(* IEC 61131-3 sources: daoli-st-library/DL_Motion (part 3) *)

(* ---- FC_DL_CamTableValidate.st ---- *)
(*
    FC_DL_CamTableValidate —— 凸轮表合法性校验
    ------------------------------------------------------------------
    分类      : DL_Motion / CamData
    前缀      : FC_DL_
    版本      : 1.0.0
    溯源      : T1-6 PLCopen MC_CamTableSelect 表选择纪律（只借「凸轮表在下装前必须
                完成相位单调、首尾闭合、斜率可行性检查」的公开语义）；
                校验算法、掩码布局、容差处理与码位 100% 自有；clean-room 重写，
                未复制任何闭源厂商源码，参考实现仅限 MIT/Apache 许可
    道莅 clean-room 防御性实现：语义借鉴、代码与码位 100% 自有
    平台      : 纯 IEC 61131-3，CODESYS V3.5+ / TwinCAT 3 / InoProShop / Machine Expert 通用
    作者      : 道莅代码库 · PLC编程专家（R22 批 4 · #15）
    ------------------------------------------------------------------
    功能说明  : 凸轮表下装前的离线校验器。一趟扫描内同时评估五项：
                ① 相位严格递增（含重复点与倒序点）② 相位值与从轴值非有限
                ③ 周期表首尾相位闭合 ④ 段斜率上限 ⑤ 有效点数合法。
                返回 TRUE = 表可用于生产（斜率超限只提示不否决）。
    不早退    : 四类判据**全部**评估完再出口，掩码一次给全——现场改一张表往往要一并
                修好几处，早退会让人改一处、重下装、再报下一处，来回好几轮。
    职责边界  : ① 只判相位闭合，不判从轴首尾等值。周期凸轮若从轴不回零点会持续漂移，
                   但这条判据不在派单掩码位内，扩位会破坏下游对掩码位含义的既有依赖；
                   建表工具必须自己保证从轴首尾等值，本函数不替它兜底。
                ② 不判表内点数以外的高阶连续性（加速度跳变、冲击），那属于工艺设计。
                ③ 不修改传入数组，纯只读。
    容差说明  : fPhaseTol 为闭合容差。容差填成负值时闭合判据必然失败（安全侧：宁可不放行），
                本函数**不钳位**——钳位会让负值变成一个「看起来正常」的容差，掩盖填表错误。
                fMaxSlope 填成非正值时任何正斜率都会触发提示码，同样按安全侧处理，不钳位。
    错误码    : 16#0004_01DB 非周期表，已跳过首尾闭合校验——信息级
                16#0004_01DC 斜率超限，表仍可用（仅提示）——信息级
                16#0004_02F3 有效点数非法 / 相位非单调（倒序或重复点）——故障级，
                             掩码位 16（点数）与位 1（单调）共用本码（R90）
                16#0004_02F4 相位值或从轴值非有限（NaN / ±Inf）——故障级，掩码位 2
                16#0004_02F5 周期表首尾相位未闭合——故障级，掩码位 4
    码位总账  : 16#0004_01DB 用 / 16#0004_01DC 用 ｜ 16#0004_02F3 用 / 16#0004_02F4 用 / 16#0004_02F5 用
    掩码总账  : 位 1 = 相位非单调（含重复点）｜ 位 2 = 相位或从轴非有限｜ 位 4 = 首尾未闭合
                ｜ 位 8 = 斜率超限｜ 位 16 = 有效点数非法｜ 其余位恒 0（预留禁用，不得挪用）
    状态机    : N/A —— 纯函数无顺序状态机，无 CASE 可写，非法状态不可能出现
    采样约定  : 纯组合函数，无定时器、无内部驻留状态，调用即出结果。
                数组按值传入（两张表各 64 × 4 字节 = 512 字节），故本函数只应在建表 /
                下装 / 参数变更事件里调用，严禁放进 1 ms 级高速循环（那是拿扫描周期换校验）。
    依赖      : 仅 Standard.library（ABS / MAX / MIN），不引用任何其他 DL_ 子库。
    验收向量  :
                V1 域外早退：uSegCount = 1 → 掩码 16#0010、uFailIdx = 0、02F3、
                   bError = TRUE、返回 FALSE。
                V2 上限/提示：表合格但某段斜率 150 mm/° > fMaxSlope 100 → 掩码 16#0008、
                   01DC、返回 TRUE、bValid = TRUE（可用但需关注）。
                V3 相位重复点：afPhase[3] = afPhase[2]（Δphase = 0）→ 掩码 16#0001、
                   uFailIdx = 3、02F3、返回 FALSE；该段不参与斜率计算（除零前置闸）。
                V4 复位/跳过首拍：bCyclic = FALSE 且其余合格 → 掩码 0、01DB、返回 TRUE。
                V5 round-trip：把同一张表分别做成「闭合的周期表（末点 = 首点 + 360°
                   且从轴末点 = 首点）」与「相位倒序的坏表」，前者 TRUE、后者 FALSE 且
                   掩码恒含位 1。
    红线自检  : 1 全局变量声明零使用 / 外部变量访问零使用 / 物理地址零使用 —— 通过，全部量经引脚传入
                2 纯 IEC 61131-3 跨平台 —— 通过，仅 Standard.library
                3 防御性编程 —— 通过，除零前置闸先判 Δphase > 0 再算商，WHILE 带 nGuard
                   计数器，数组索引全部由已校验的点数上限约束
                4 声明行同行中英双语注释 + 单位 —— 通过，逐行附注
                5 ENUM + CASE —— 不适用（纯函数，状态机 N/A，头注释已声明）
                6 TON / R_TRIG —— 不适用（无实例、无周期驻留）
                7 无魔法数 —— 通过，点数上下限、掩码位、整圈角度全部 VAR CONSTANT
    修订记录  : 2026-11-16 v1.0.0 首次入库（R22 批 4 · #15）
*)
FUNCTION FC_DL_CamTableValidate : BOOL
VAR_INPUT
    afPhase     : ARRAY[0..DL_CAM_LAST_IDX] OF REAL;   // 相位表 [°]，须严格递增 / phase table [deg], must strictly increase
    afSlave     : ARRAY[0..DL_CAM_LAST_IDX] OF REAL;   // 从轴位置表 [mm]，与相位表同下标 / slave position table [mm], indexed like the phase table
    uSegCount   : UINT := 8;                   // 有效点数 [个]，范围 2~64 / number of valid points [pcs], range 2..64
    bCyclic     : BOOL := TRUE;                // 周期表须首尾相位闭合 / a cyclic table must close its phase across the wrap
    fPhaseTol   : REAL := 0.01;                // 闭合容差 [°]，负值即判闭合失败 / closure tolerance [deg], a negative value fails the check
    fMaxSlope   : REAL := 100.0;               // 段斜率上限 [mm/°]，仅提示不否决 / segment slope limit [mm/deg], informational only
END_VAR
VAR_OUTPUT
    uFailMask      : WORD;                     // 失败掩码，全部失败项同时置位 / failure mask, every failing criterion is set at once
    uFailIdx       : UINT;                     // 1 基首个失败段号，0 = 无 / one-based index of the first failing segment, 0 = none
    fMaxSlopeFound : REAL;                     // 实测最大段斜率 [mm/°] / largest measured segment slope [mm/deg]
    eErr           : UDINT;                    // 错误码，0 表示无错 / error code, 0 means no error
    bError         : BOOL;                     // 故障级标志，仅故障级错误置位 / fault-class flag, set only on fault-level codes
    bValid         : BOOL;                     // 校验结论可信标志，= NOT bError / verdict trustworthy flag, equals NOT bError
END_VAR
VAR
    uSegUse     : UINT;                        // 校验时实际使用的点数，已过范围门禁 / point count actually used after the range gate
    uMaskWork   : WORD;                        // 掩码累加器，出口一次性发布 / mask accumulator published once at the exit
    uIdxWork    : UINT;                        // 首个失败段号累加器 / first failing segment accumulator
    nI          : UINT;                        // 扫描下标 [个] / scan index [pcs]
    nGuard      : UINT;                        // 循环保护计数器，上限 DL_CAM_GUARD / loop guard counter bounded by DL_CAM_GUARD
    fDp         : REAL;                        // 本段相位增量 [°] / phase increment of this segment [deg]
    fDs         : REAL;                        // 本段从轴增量 [mm] / slave increment of this segment [mm]
    fSlope      : REAL;                        // 本段斜率 [mm/°] / slope of this segment [mm/deg]
    fClose      : REAL;                        // 首尾相位闭合偏差（已减整圈）[°] / closure deviation after removing one full turn [deg]
END_VAR
VAR CONSTANT
    DL_CAM_LAST_IDX  : UINT := 63;             // 数组末下标 [下标]，即点数上限 64 / last array index, i.e. a capacity of 64 points
    DL_CAM_SEG_MIN   : UINT := 2;              // 有效点数下限 [个] / lower bound of the point count [pcs]
    DL_CAM_SEG_MAX   : UINT := 64;             // 有效点数上限 [个] / upper bound of the point count [pcs]
    DL_CAM_GUARD     : UINT := 64;             // 循环保护上限 [拍]，与点数上限同源 / loop guard bound [scans], tied to the point capacity
    DL_CAM_FULL_TURN : REAL := 360.0;          // 整圈角度 [°] / one full turn [deg]
    DL_CAM_ZERO      : REAL := 0.0;            // 零值常量，避免裸字面量 [无量纲] / zero constant, avoids a bare literal [dimensionless]
    DL_CAM_MK_MONO   : WORD := 16#0001;        // 掩码位 1：相位非单调（含重复点）/ mask bit 1, the phase is not increasing
    DL_CAM_MK_FIN    : WORD := 16#0002;        // 掩码位 2：相位或从轴非有限 / mask bit 2, a phase or slave value is not finite
    DL_CAM_MK_CLOSE  : WORD := 16#0004;        // 掩码位 4：首尾相位未闭合 / mask bit 4, the phase does not close
    DL_CAM_MK_SLOPE  : WORD := 16#0008;        // 掩码位 8：斜率超限（仅提示）/ mask bit 8, the slope exceeds the limit, informational
    DL_CAM_MK_COUNT  : WORD := 16#0010;        // 掩码位 16：有效点数非法 / mask bit 16, the point count is illegal
    DL_CAM_MK_NONE   : WORD := 16#0000;        // 空掩码常量，避免裸字面量比较 / empty mask constant, avoids a bare literal comparison
END_VAR

// 段 1｜预置：掩码与段号先清零，出口一次性发布（R94 统一后处理）
// segment 1, preset the mask and the index so the exit publishes them once
uMaskWork := DL_CAM_MK_NONE;                    // 掩码清零 / clear the mask
uIdxWork := 0;                                  // 段号清零，0 = 无失败 / clear the index, 0 = none
fMaxSlopeFound := DL_CAM_ZERO;                  // 实测斜率清零 / clear the measured slope
eErr := 0;                                      // 预置无错误 / preset no error
bError := FALSE;                                // 预置无故障标志 / preset no error flag

// 段 2｜点数门禁：点数非法时后面任何判据都无从谈起，这是唯一的例外早退
// segment 2, the point-count gate, the only early exit because no criterion can be evaluated without a legal count
IF (uSegCount < DL_CAM_SEG_MIN) OR (uSegCount > DL_CAM_SEG_MAX) THEN
    uMaskWork := uMaskWork OR DL_CAM_MK_COUNT;  // 掩码位 16：有效点数非法 / mask bit 16, illegal point count
    uIdxWork := 0;                              // 点数非法时没有「失败段」可言 / an illegal count has no failing segment
    uFailMask := uMaskWork;                     // 发布掩码 / publish the mask
    uFailIdx := uIdxWork;                       // 发布段号 / publish the index
    fMaxSlopeFound := DL_CAM_ZERO;              // 未做扫描，斜率无实测值 / no scan was run so there is no measured slope
    eErr := 16#0004_02F3;                       // 故障级：点数非法（与单调失败共用本码，R90）/ fault: illegal count, shared with the monotonic failure
    bError := TRUE;                             // 置故障标志 / raise the fault flag
    bValid := FALSE;                            // 结论不可信 / the verdict is not trustworthy
    FC_DL_CamTableValidate := FALSE;            // 表不可用 / the table is not usable
ELSE
    uSegUse := uSegCount;                       // 点数合法，按实际点数扫描 / a legal count, scan the actual point set

    // 段 3｜单趟扫描：非有限检测与相位单调/斜率同环评估，绝不早退（R94 掩码要全）
    // segment 3, one pass evaluating the finiteness and the monotonic/slope criteria together, never exiting early
    nI := 0;                                    // 下标起点 / start the index at zero
    nGuard := 0;                                // 循环保护计数清零 / clear the loop guard
    WHILE (nI < uSegUse) AND (nGuard < DL_CAM_GUARD) DO
        // 3.1 非有限检测：同一式兼捕 NaN 与 ±Inf —— Inf 减 Inf 得 NaN，故自不自等同样成立；
        //     有限值减自身恒为 0，不会误报。
        // non-finite detection, one test catches NaN and plus/minus infinity alike while a finite value subtracts to zero
        IF (afSlave[nI] - afSlave[nI]) <> (afSlave[nI] - afSlave[nI]) THEN
            uMaskWork := uMaskWork OR DL_CAM_MK_FIN;    // 从轴值非有限 / the slave value is not finite
            IF uIdxWork = 0 THEN
                IF nI > 0 THEN
                    uIdxWork := nI;             // 该点所在段的段号（1 基）/ the segment that ends at this point
                ELSE
                    uIdxWork := 1;              // 首点归属第 1 段 / the first point belongs to segment one
                END_IF
            END_IF
        END_IF
        IF (afPhase[nI] - afPhase[nI]) <> (afPhase[nI] - afPhase[nI]) THEN
            uMaskWork := uMaskWork OR DL_CAM_MK_FIN;    // 相位值非有限，与从轴共用掩码位 2 / a non-finite phase shares mask bit 2
            IF uIdxWork = 0 THEN
                IF nI > 0 THEN
                    uIdxWork := nI;             // 该点所在段的段号（1 基）/ the segment that ends at this point
                ELSE
                    uIdxWork := 1;              // 首点归属第 1 段 / the first point belongs to segment one
                END_IF
            END_IF
        END_IF

        // 3.2 相位单调与段斜率：增量非正一律判单调失败，且绝不进入除法（除零前置闸）
        // monotonic test and slope, a non-positive increment fails the criterion and never reaches the division
        IF nI > 0 THEN
            fDp := afPhase[nI] - afPhase[nI - 1];   // 本段相位增量 [°] / phase increment of this segment [deg]
            IF NOT (fDp > DL_CAM_ZERO) THEN         // 含 0（重复点）、负（倒序）与 NaN 三种情形 / covers a duplicate, a reversal and NaN alike
                uMaskWork := uMaskWork OR DL_CAM_MK_MONO;   // 掩码位 1：相位非单调 / mask bit 1, the phase is not increasing
                IF uIdxWork = 0 THEN
                    uIdxWork := nI;             // 失败段号 = 末点序号（1 基）/ the failing segment equals the ending point index
                END_IF
            ELSE
                fDs := afSlave[nI] - afSlave[nI - 1];   // 本段从轴增量 [mm] / slave increment of this segment [mm]
                fSlope := ABS(fDs / fDp);               // 斜率绝对值，除子已判正 [mm/°] / absolute slope with a guarded divisor [mm/deg]
                IF fSlope > fMaxSlopeFound THEN
                    fMaxSlopeFound := fSlope;           // 记录实测最大斜率 / keep the largest measured slope
                END_IF
            END_IF
        END_IF

        nI := nI + 1;                           // 下标推进 / advance the index
        nGuard := nGuard + 1;                   // 保护计数推进 / advance the guard
    END_WHILE

    // 段 4｜首尾闭合：仅周期表判，非周期表跳过并留信息码
    // segment 4, closure check applied to cyclic tables only, a non-cyclic table skips it and leaves an info code
    IF bCyclic THEN
        fClose := afPhase[uSegUse - 1] - afPhase[0] - DL_CAM_FULL_TURN;     // 闭合偏差已去掉整圈 [°] / deviation after removing one full turn [deg]
        IF ABS(fClose) > fPhaseTol THEN
            uMaskWork := uMaskWork OR DL_CAM_MK_CLOSE;   // 掩码位 4：首尾相位未闭合 / mask bit 4, the phase does not close
            IF uIdxWork = 0 THEN
                uIdxWork := uSegUse;        // 闭合段是第 N 段（末点回到首点）/ the wrap segment is segment N, the last point back to the first
            END_IF
        END_IF
    END_IF

    // 段 5｜斜率提示：超限只置掩码位 8，绝不否决表（工艺上宽斜率常是有意为之）
    // segment 5, the slope hint sets mask bit 8 only, a wide slope is often deliberate and never rejects the table
    IF (fMaxSlopeFound > fMaxSlope) THEN
        uMaskWork := uMaskWork OR DL_CAM_MK_SLOPE;  // 掩码位 8：斜率超限（仅提示）/ mask bit 8, the slope exceeds the limit, informational only
    END_IF

    // 段 6｜错误码优先级：故障码先占，其次斜率提示，最后非周期提示（同拍只发一条，R45）
    // segment 6, code priority, faults first then the slope hint then the non-cyclic notice, one code per scan
    IF (uMaskWork AND DL_CAM_MK_MONO) <> DL_CAM_MK_NONE THEN
        eErr := 16#0004_02F3;                   // 故障级：相位非单调或点数非法（共用本码，R90）/ fault: the phase is not increasing or the count is illegal, shared code
        bError := TRUE;
    ELSIF (uMaskWork AND DL_CAM_MK_FIN) <> DL_CAM_MK_NONE THEN
        eErr := 16#0004_02F4;                   // 故障级：相位或从轴非有限 / fault: a phase or slave value is not finite
        bError := TRUE;
    ELSIF (uMaskWork AND DL_CAM_MK_CLOSE) <> DL_CAM_MK_NONE THEN
        eErr := 16#0004_02F5;                   // 故障级：周期表首尾相位未闭合 / fault: the cyclic table does not close
        bError := TRUE;
    ELSIF (uMaskWork AND DL_CAM_MK_SLOPE) <> DL_CAM_MK_NONE THEN
        eErr := 16#0004_01DC;                   // 信息级：斜率超限，表仍可用 / info: the slope exceeds the limit and the table stays usable
    ELSIF NOT bCyclic THEN
        eErr := 16#0004_01DB;                   // 信息级：非周期表，已跳过闭合校验 / info: a non-cyclic table skipped the closure check
    END_IF

    // 段 7｜出口：掩码与段号一次性发布，返回可用性
    // segment 7, publish the mask and the index once and return the usability
    uFailMask := uMaskWork;                     // 发布掩码（全部失败项同时给全）/ publish the mask with every failing criterion
    uFailIdx := uIdxWork;                       // 发布首个失败段号 / publish the first failing segment
    bValid := NOT bError;                       // 结论可信 = 无故障级错误（斜率提示不影响可信）/ the verdict is trustworthy without a fault-level code
    FC_DL_CamTableValidate := NOT bError;       // 返回 TRUE = 表可用 / TRUE means the table is usable
END_IF
END_FUNCTION

(* ---- FC_DL_ChainWearElongation.st ---- *)
(*
  ============================================================
  组件名 : FC_DL_ChainWearElongation
  分类   : DL_Motion
  功能   : 链条磨损伸长率计算，由公称节距与实测节距求伸长百分比并给出更换到期判定
  复杂度 : C1
  版本   : 1.0.0
  作者   : 道莅工业代码库工厂 / R81
  日期   : 2026-11-24
  开源溯源 : clean-room（no upstream）—— 依据公开工程公式自研，未复制任何上游实现
  红线自检 : R1 无GVL/R2 无物理地址/R3 纯IEC/R4 防除零/R5 双语注释
  接口说明 :
      伸长率 = (实测节距 - 公称节距) / 公称节距 * 100。
      实测节距必须为多节平均后的值，节数少于 3 节时平均值不具代表性，判无效。
      伸长率超过 2.0% 判更换到期；实测小于公称（新链或测量误差）时伸长率为负，判定位保持 FALSE。
  ============================================================
*)
FUNCTION FC_DL_ChainWearElongation : BOOL
VAR_INPUT
    bEnable      : BOOL; // 使能：TRUE 时计算 / Enable: TRUE to compute
    bErr         : BOOL; // 外部故障：TRUE 时立即退出并置结果无效 / External fault: TRUE aborts with invalid result
    rPitchNom_mm : REAL; // 公称节距 [mm] / nominal chain pitch [millimetre]
    rPitchAct_mm : REAL; // 实测节距，取多节平均 [mm] / measured pitch averaged over several links [millimetre]
    iLinkCnt     : INT;  // 参与平均的链节数量 [节] / number of links used in the average [link]
END_VAR
VAR_OUTPUT
    rElongPct   : REAL; // 链条磨损伸长率 [%] / chain wear elongation [percent]
    rPitchDelta_mm : REAL; // 实测与公称的节距差 [mm] / pitch difference between the measured and nominal value [millimetre]
    bReplaceDue : BOOL; // 更换到期：TRUE 表示伸长率超过 2.0% / replacement due, TRUE when the elongation exceeds 2.0 percent
    bValid      : BOOL; // 输出有效：TRUE 表示结果可用 / Output valid
END_VAR
VAR CONSTANT
    DL_R_MAX    : REAL := 3.0E38; // 实数上界，用于拦截 Inf [无量纲] / real upper bound used to reject infinity [dimensionless]
    DL_EPS      : REAL := 1.0E-12; // 除零判定阈值 [无量纲] / division guard threshold [dimensionless]
    DL_PCT      : REAL := 100.0;  // 百分数换算系数 [无量纲] / percentage scaling factor [dimensionless]
    DL_ELONG_MAX : REAL := 2.0;   // 更换到期伸长率门限 [%] / elongation threshold for the replacement [percent]
    DL_LINK_MIN : INT := 3;       // 平均所需最少链节数 [节] / minimum link count required by the average [link]
    DL_LINK_MAX : INT := 200;     // 链节数量合理上限 [节] / sanity upper bound of the link count [link]
    DL_PITCH_MAX : REAL := 1000.0; // 节距合理上限 [mm] / sanity upper bound of the pitch [millimetre]
END_VAR
VAR
    _bFin : BOOL := FALSE; // 输入有限性判定结果 / input finiteness verdict
END_VAR

    // 段 1｜出口预置
    rElongPct := 0.0;
    rPitchDelta_mm := 0.0;
    bReplaceDue := FALSE;
    bValid := FALSE;
    // 段 2｜使能闸与外部故障闸
    IF NOT bEnable THEN
        RETURN;
    END_IF;
    IF bErr THEN
        RETURN;
    END_IF;
    // 段 3｜非有限闸
    _bFin := (rPitchNom_mm = rPitchNom_mm) AND (ABS(rPitchNom_mm) <= DL_R_MAX) AND (rPitchAct_mm = rPitchAct_mm) AND (ABS(rPitchAct_mm) <= DL_R_MAX);
    IF NOT _bFin THEN
        RETURN;
    END_IF;
    // 段 4｜域闸：公称节距严格为正且合理，实测节距非负且合理，链节数 3~200
    IF (ABS(rPitchNom_mm) <= DL_EPS) OR (rPitchNom_mm < 0.0) OR (rPitchNom_mm > DL_PITCH_MAX) THEN
        RETURN;
    END_IF;
    IF (rPitchAct_mm < 0.0) OR (rPitchAct_mm > DL_PITCH_MAX) THEN
        RETURN;
    END_IF;
    IF (iLinkCnt < DL_LINK_MIN) OR (iLinkCnt > DL_LINK_MAX) THEN
        RETURN;
    END_IF;
    // 段 5｜节距差与伸长率
    rPitchDelta_mm := rPitchAct_mm - rPitchNom_mm;
    rElongPct := rPitchDelta_mm / rPitchNom_mm * DL_PCT;
    // 段 6｜更换到期判定：仅正向伸长计入磨损
    IF rElongPct > DL_ELONG_MAX THEN
        bReplaceDue := TRUE;
    ELSE
        bReplaceDue := FALSE;
    END_IF;
    bValid := TRUE;
    FC_DL_ChainWearElongation := bValid;
END_FUNCTION

(* ---- FC_DL_CornerRoundingRadiusCalc.st ---- *)
(* ============================================================
   DL_Motion / FC_DL_CornerRoundingRadiusCalc ｜ v1.0.0 ｜ 2026-11-25
   功能：拐角圆弧过渡半径 [mm] 与拐角通过速度 [mm/min]：
         r ≤ min(段长)/2 × tan(θ/2)（切线长约束，另受 20 mm 工艺硬上限）；
         v ≤ (j·r²)^(1/3)（jerk 约束，再与编程进给取小）
   边界：θ∉(0,180)° / 段长≤0 / 进给≤0 / jerk≤0 或非有限 → 半径与速度写 0（N1/N3）；
         fJerkRatio = v_use³/(r²·j) ∈ [0,1]，v_use = 实际采用进给（mm/s），
         = 1 表示 jerk 用满、< 1 表示受编程进给限制（N5 系数回代）
   依赖：仅 IEC 61131-3（SQRT / EXPT / TAN / MIN） ｜ 溯源：DLF-A-RTCP（内部原创线）
   ============================================================ *)
FUNCTION FC_DL_CornerRoundingRadiusCalc : BOOL
VAR_INPUT
    fCornerAngleDeg : LREAL;  // 拐角夹角，域 (0,180) [deg] / Corner included angle
    fSegLenAMm      : LREAL;  // 前一段长度，域 > 0 [mm] / Length of the incoming segment
    fSegLenBMm      : LREAL;  // 后一段长度，域 > 0 [mm] / Length of the outgoing segment
    fFeedMaxMmMin   : LREAL;  // 编程进给上限，域 > 0 [mm/min] / Programmed feed ceiling
    fJerkMaxMmS3    : LREAL;  // 允许 jerk 上限，域 > 0 [mm/s³] / Allowed jerk ceiling
END_VAR
VAR_OUTPUT
    fRadiusMm        : LREAL;  // 过渡圆弧半径 [mm] / Rounding arc radius
    fCornerFeedMmMin : LREAL;  // 拐角通过速度 [mm/min] / Corner pass-through feed rate
    fJerkRatio       : REAL;   // jerk 使用率 [0,1] [-] / Jerk utilization ratio
END_VAR
VAR
    _fThetaRad : LREAL;  // 夹角弧度值 [rad] / Included angle in radians
    _fRmax     : LREAL;  // 段长约束下的半径上限 [mm] / Radius ceiling from segment lengths
    _fVuse     : LREAL;  // jerk 约束允许速度 [mm/s] / Speed allowed by the jerk limit
    _fVact     : LREAL;  // 实际采用进给（换算到 mm/s）[mm/s] / Adopted feed rate in millimeters per second
END_VAR
VAR CONSTANT
    DL_CRN_PI : LREAL := 3.14159265358979324;  // 圆周率（LREAL 全精度）[-] / Pi at full precision
END_VAR

(* 段 0：出口预置安全侧（半径 0 = 不做过渡，N3） *)
FC_DL_CornerRoundingRadiusCalc := FALSE;
fRadiusMm := 0.0;  fCornerFeedMmMin := 0.0;  fJerkRatio := 0.0;

(* 段 1：非有限闸 + 五域闸（夹角开区间、四个正值域） *)
IF (fCornerAngleDeg <> fCornerAngleDeg) OR (fSegLenAMm <> fSegLenAMm)
   OR (fSegLenBMm <> fSegLenBMm) OR (fFeedMaxMmMin <> fFeedMaxMmMin)
   OR (fJerkMaxMmS3 <> fJerkMaxMmS3) THEN
    RETURN;
END_IF
IF (fCornerAngleDeg <= 0.0) OR (fCornerAngleDeg >= 180.0) THEN RETURN; END_IF
IF (fSegLenAMm <= 0.0) OR (fSegLenBMm <= 0.0) THEN RETURN; END_IF
IF (fFeedMaxMmMin <= 0.0) OR (fJerkMaxMmS3 <= 0.0) THEN RETURN; END_IF

(* 段 2：半径上限（切线长 T = r/tan(θ/2) ≤ 最短段长/2）与硬上限 *)
_fThetaRad := fCornerAngleDeg * DL_CRN_PI / 180.0;
_fRmax := (MIN(fSegLenAMm, fSegLenBMm) / 2.0) * TAN(_fThetaRad / 2.0);
fRadiusMm := MIN(_fRmax, 20.0);                          // 20 mm 工艺硬上限

(* 段 3：jerk 约束速度 v = (j·r²)^(1/3) [mm/s]，再与编程进给取小 *)
_fVuse := EXPT(fJerkMaxMmS3 * fRadiusMm * fRadiusMm, 0.33333333333333333);
fCornerFeedMmMin := MIN(fFeedMaxMmMin, _fVuse * 60.0);   // mm/s → mm/min

(* 段 4：jerk 使用率（按实际采用进给回代：v_use = fCornerFeedMmMin/60；
   代 _fVuse 回代会代数恒等为 1.000000，输出无信息量，故改用采用值） *)
_fVact := fCornerFeedMmMin / 60.0;                       // mm/min → mm/s
fJerkRatio := LREAL_TO_REAL((_fVact * _fVact * _fVact) / (fRadiusMm * fRadiusMm * fJerkMaxMmS3));
IF (fJerkRatio <> fJerkRatio) OR ((fJerkRatio - fJerkRatio) <> (fJerkRatio - fJerkRatio))
   OR (fJerkRatio < 0.0) THEN fJerkRatio := 0.0; END_IF
IF fJerkRatio > 1.0 THEN fJerkRatio := 1.0; END_IF

(* 段 5：结果复检 + 单一出口裁决（N4） *)
IF (fRadiusMm <> fRadiusMm) OR ((fRadiusMm - fRadiusMm) <> (fRadiusMm - fRadiusMm))
   OR (fCornerFeedMmMin <> fCornerFeedMmMin)
   OR ((fCornerFeedMmMin - fCornerFeedMmMin) <> (fCornerFeedMmMin - fCornerFeedMmMin)) THEN
    fRadiusMm := 0.0;  fCornerFeedMmMin := 0.0;  fJerkRatio := 0.0;  RETURN;
END_IF
FC_DL_CornerRoundingRadiusCalc := TRUE;
END_FUNCTION

(* ---- FC_DL_DiffDriveOdometryCalc.st ---- *)
// FC_DL_DiffDriveOdometryCalc v1.0.0
// 开源溯源：clean-room 自研（族 DL_Motion，ST 生态实测 0 命中，无外部代码引入）
(*
  功能: 差速轮单周期里程计：ds = (dR+dL)/2，dθ = (dR−dL)/B，
        dx = ds·COS(θ + dθ/2)，dy = ds·SIN(θ + dθ/2)，θnew = θ + dθ 归一化到 (−π, π]。
  邻件/码位: 为路径跟踪链的定位侧件（只产生位姿增量，不含跟踪律）；
             16#0002_9203 = 域外、非有限或归一化不收敛拒收。
*)
FUNCTION FC_DL_DiffDriveOdometryCalc : REAL
VAR_INPUT
    fDeltaLeft  : REAL := 0.0;      // 左轮增量位移 [m]，前进正 / Left incremental travel [m]
    fDeltaRight : REAL := 0.0;      // 右轮增量位移 [m]，前进正 / Right incremental travel [m]
    fWheelBase  : REAL := 0.5;      // 轮距 B [m]，域 > 1e-6 / Wheel base [m]
    fThetaPrev  : REAL := 0.0;      // 上周期航向 θ [rad] / Previous heading [rad]
END_VAR
VAR_OUTPUT
    fDeltaX   : REAL;               // 本周期 X 增量 [m] / Incremental X displacement [m]
    fDeltaY   : REAL;               // 本周期 Y 增量 [m] / Incremental Y displacement [m]
    fThetaNew : REAL;               // 归一化新航向 (−π, π] [rad] / Normalized heading [rad]
    fDeltaS   : REAL;               // 本周期弧长增量 [m] / Incremental arc length [m]
    bValid    : BOOL;               // 结果有效回执 [-] / Result validity receipt
    uErrorId  : UDINT;              // 事件码，0 = 无事件 / Event code
END_VAR
VAR
    fPi    : REAL := 3.14159265358979;  // 圆周率常量 [rad] / Pi constant [rad]
    fTwoPi : REAL := 6.28318530717959;  // 二倍圆周率 [rad] / Two pi constant [rad]
    fDTheta : REAL := 0.0;          // 本周期航向增量 dθ [rad] / Heading increment [rad]
    iGuard : INT := 0;              // 归一化循环守卫计数 [次] / Normalization loop guard
END_VAR
// 段 0：全路径出口安全缺省（航向回绝对零，不回灌上拍）/ Safe defaults, heading to absolute zero
fDeltaX := 0.0;                     // X 增量缺省零 / X increment default zero
fDeltaY := 0.0;                     // Y 增量缺省零 / Y increment default zero
fDeltaS := 0.0;                     // 弧长增量缺省零 / Arc increment default zero
fThetaNew := 0.0;                   // 航向缺省绝对零 / Heading default absolute zero
bValid := FALSE;                    // 有效回执预清 / Validity preset clear
uErrorId := 16#0000;                // 事件码预清 / Event code preset clear
FC_DL_DiffDriveOdometryCalc := 0.0; // 返回值缺省零（镜像弧长）/ Return default zero
// 段 1：非有限闸（四入参全枚举）/ Non-finite gate over all inputs
IF (fDeltaLeft <> fDeltaLeft) OR (fDeltaRight <> fDeltaRight)
   OR (fWheelBase <> fWheelBase) OR (fThetaPrev <> fThetaPrev)
   OR (ABS(fDeltaLeft) >= 3.0E38) OR (ABS(fDeltaRight) >= 3.0E38)
   OR (ABS(fWheelBase) >= 3.0E38) OR (ABS(fThetaPrev) >= 3.0E38) THEN
    uErrorId := 16#0002_9203;   // 入参非有限拒收 / Non-finite input reject
    RETURN;
END_IF
// 段 2：域闸（轮距为正，dθ 分母非零）/ Domain gate, R4 divide-by-zero guard
IF fWheelBase <= 1.0E-6 THEN
    uErrorId := 16#0002_9203;   // 轮距非正，航向不可解 / Non-positive wheel base
    RETURN;
END_IF
// 段 3：主计算（中点积分 + 航向归一化）/ Main computation with heading normalization
fDeltaS := (fDeltaRight + fDeltaLeft) / 2.0;                    // 弧长增量 / Arc increment
fDTheta := (fDeltaRight - fDeltaLeft) / fWheelBase;             // 航向增量 / Heading increment
fDeltaX := fDeltaS * COS(fThetaPrev + fDTheta / 2.0);           // X 增量（半角）/ X increment half-angle
fDeltaY := fDeltaS * SIN(fThetaPrev + fDTheta / 2.0);           // Y 增量（半角）/ Y increment half-angle
fThetaNew := fThetaPrev + fDTheta;                              // 未归一化航向 / Raw new heading
iGuard := 0;                                                    // 守卫计数清零 / Guard counter clear
WHILE (fThetaNew > fPi) AND (iGuard < 64) DO                    // 超上界折叠 / Fold above upper bound
    fThetaNew := fThetaNew - fTwoPi;                            // 减一整周 / Subtract one turn
    iGuard := iGuard + 1;                                       // 守卫自增 / Guard increment
END_WHILE
WHILE (fThetaNew <= -fPi) AND (iGuard < 64) DO                  // 超下界折叠 / Fold below lower bound
    fThetaNew := fThetaNew + fTwoPi;                            // 加一整周 / Add one turn
    iGuard := iGuard + 1;                                       // 守卫自增 / Guard increment
END_WHILE
// 段 4：出口闸（非有限复核 + 归一化收敛复核）/ Outlet gate
IF (fDeltaX <> fDeltaX) OR (fDeltaY <> fDeltaY) OR (fDeltaS <> fDeltaS) OR (fThetaNew <> fThetaNew)
   OR (ABS(fDeltaX) >= 3.0E38) OR (ABS(fDeltaY) >= 3.0E38)
   OR (ABS(fDeltaS) >= 3.0E38) OR (ABS(fThetaNew) >= 3.0E38) THEN
    fDeltaX := 0.0;             // 复核失败回缺省 / Fallback on recheck failure
    fDeltaY := 0.0;             // 复核失败回缺省 / Fallback on recheck failure
    fDeltaS := 0.0;             // 复核失败回缺省 / Fallback on recheck failure
    fThetaNew := 0.0;           // 复核失败回绝对零 / Heading falls back to absolute zero
    uErrorId := 16#0002_9203;   // 出口非有限拒收 / Output non-finite reject
    RETURN;
END_IF
IF iGuard >= 64 THEN
    uErrorId := 16#0002_9203;   // 归一化未收敛（航向超 64 周）/ Normalization not converged
    RETURN;
END_IF
bValid := TRUE;                 // 有效回执 / Validity receipt
FC_DL_DiffDriveOdometryCalc := fDeltaS;     // 返回值镜像弧长增量 / Return mirrors arc increment
END_FUNCTION

(* ---- FC_DL_GearRatioCalc.st ---- *)
// FC_DL_GearRatioCalc v1.0.0
// 开源溯源：self-cleanroom / 机械传动族
(*
  道莅工业代码库 | DL_Motion | FC_DL_GearRatioCalc
  版本: 1.0.0 | 日期: 2026-11-23 | 轮次: R75
  功能: 齿轮减速比与负载惯量比换算：减速比 i = n_in/n_out = z_out/z_in，
        折算负载惯量 J_ref = J_load / i²（负载侧经减速机折算至电机侧）
  邻件关系: 与 GearInPhaseAlign（齿轮相位对齐）同族 —— 差异点：相位件做
            啮合相位对齐动作，本件为纯比值/折算计算件，无相位语义；
            本件码位 16#0002_2601
*)
FUNCTION FC_DL_GearRatioCalc : REAL
VAR_INPUT
    fSpeedIn   : REAL := 0.0;   // 输入转速 n_in [rpm]，域 > 0 / Input speed [rpm], domain > 0
    fSpeedOut  : REAL := 0.0;   // 输出转速 n_out [rpm]，域 > 0 / Output speed [rpm], domain > 0
    fLoadInertia: REAL := 0.0;  // 负载侧惯量 J_load [kg·m²]，域 >= 0 / Load-side inertia [kg·m2]
    fEps       : REAL := 1.0E-6;// 判零容差 [rpm|kg·m²] / Zero tolerance
END_VAR
VAR_OUTPUT
    fRatio     : REAL;          // 减速比 i = n_in/n_out [1] / Gear ratio
    fInertiaRef: REAL;          // 折算至电机侧负载惯量 J_load/i² [kg·m²] / Load inertia referred to motor side
    bValid     : BOOL;          // 结果有效回执 [-] / Result validity receipt
    uErrorId   : UDINT;         // 事件码，0 = 无事件；16#0002_2601 = 域外拒收 / Event code
END_VAR

// —— 段 0：全路径缺省 —— //
fRatio := 0.0;                   // 减速比缺省零 / Ratio default zero
fInertiaRef := 0.0;              // 折算惯量缺省零 / Referred inertia default zero
bValid := FALSE;                 // 有效回执预清 / Validity preset
uErrorId := 16#0000;             // 事件码预清 / Event code preset
FC_DL_GearRatioCalc := 0.0;      // 返回值缺省零（镜像减速比）/ Return default mirrors ratio

// —— 段 1：非有限闸 —— //
IF (fSpeedIn <> fSpeedIn) OR (fSpeedOut <> fSpeedOut) OR (fLoadInertia <> fLoadInertia)
   OR (ABS(fSpeedIn) >= 3.0E38) OR (ABS(fSpeedOut) >= 3.0E38) OR (ABS(fLoadInertia) >= 3.0E38) THEN
    uErrorId := 16#0002_2601;    // 输入非有限拒收 / Non-finite reject
    RETURN;
END_IF

// —— 段 2：分母防零与域闸（R4） —— //
IF (fSpeedOut < fEps) OR (fSpeedIn < fEps) OR (fLoadInertia < 0.0) THEN
    uErrorId := 16#0002_2601;    // 信息级：转速非正（分母为零风险）或惯量为负 / Info level: nonpositive speed or negative inertia
    RETURN;                      // 不计算返回 / Return without computation
END_IF

// —— 段 3：主计算（分母已过闸） —— //
fRatio := fSpeedIn / fSpeedOut;  // 减速比 i = n_in/n_out / Ratio
IF fRatio < fEps THEN
    uErrorId := 16#0002_2601;    // 信息级：减速比退化近零（疑输入颠倒）/ Info level: degenerate ratio
    RETURN;
END_IF
fInertiaRef := fLoadInertia / (fRatio * fRatio);   // 折算惯量 J_load/i²（i² 非零已过闸）/ Referred inertia
bValid := TRUE;                  // 有效回执 / Validity receipt
FC_DL_GearRatioCalc := fRatio;   // 返回值 = 减速比 / Return equals ratio
END_FUNCTION

(* ---- FC_DL_HelicalTurnAdvanceCalc.st ---- *)
(* ============================================================
   DL_Motion / FC_DL_HelicalTurnAdvanceCalc ｜ v1.0.0 ｜ 2026-11-25
   功能：螺旋插补每转 Z 向进给 [mm/rev] 与切向合成进给 [mm/min]：
         合成 = √(切向² + (螺距×转速)²)，并用每转弧长 2πR 校验升角。
   边界：螺距≤0/半径≤0/转速≤0 → 码 1/2/3；非有限 → 码 4（实值同步写 0，N1）；
         螺距 > 2πR（升角>45°，自锁性丧失）→ 码 5，值照给但返回 FALSE。
   依赖：仅 IEC 61131-3（SQRT） ｜ 溯源：DLF-A-RTCP（内部原创线）
   ============================================================ *)
FUNCTION FC_DL_HelicalTurnAdvanceCalc : BOOL
VAR_INPUT
    fPitchMmRev    : LREAL;  // 螺距即每转 Z 进给，域 > 0 [mm/rev] / Helical pitch per revolution
    fRadiusMm      : LREAL;  // 螺旋中心线半径，域 > 0 [mm] / Helical centerline radius
    fFeedProgMmMin : LREAL;  // 编程切向进给率，域 > 0 [mm/min] / Programmed tangential feed rate
    fSpindleRpm    : REAL;   // 主轴转速，域 > 0 [r/min] / Spindle speed per minute
END_VAR
VAR_OUTPUT
    fZPerRev        : REAL;   // 每转 Z 向进给（等于螺距）[mm/rev] / Z advance per revolution
    fHelixFeedMmMin : REAL;   // 切向合成进给率 [mm/min] / Resulting helical feed rate
    uErrId          : UDINT;  // 出口码 0/1/2/3/4/5 [-] / Outlet code
END_VAR
VAR
    _fRpS       : LREAL;  // 转速实数值 [r/min] / Spindle speed as a real number
    _fArcPerRev : LREAL;  // 每转弧长 2πR [mm/rev] / Arc length per revolution
    _fVzMmMin   : LREAL;  // 轴向速率 = 螺距×转速 [mm/min] / Axial velocity from pitch times speed
    _fSumSq     : LREAL;  // 合成平方和 [mm²/min²] / Sum of squared velocity components
    _uCode      : UDINT;  // 出口码暂存 [-] / Staged outlet code
END_VAR
VAR CONSTANT
    DL_HEL_PI : LREAL := 3.14159265358979324;  // 圆周率（LREAL 全精度）[-] / Pi at full precision
END_VAR

(* 段 0：出口预置安全侧 *)
FC_DL_HelicalTurnAdvanceCalc := FALSE;
fZPerRev := 0.0;  fHelixFeedMmMin := 0.0;  uErrId := 4;

(* 段 1：非有限闸 + 三域闸（防零） *)
IF (fPitchMmRev <> fPitchMmRev) OR (fRadiusMm <> fRadiusMm)
   OR (fFeedProgMmMin <> fFeedProgMmMin) OR (fSpindleRpm <> fSpindleRpm) THEN
    RETURN;
END_IF
IF fPitchMmRev <= 0.0 THEN uErrId := 1; RETURN; END_IF
IF fRadiusMm <= 0.0 THEN uErrId := 2; RETURN; END_IF
IF fSpindleRpm <= 0.0 THEN uErrId := 3; RETURN; END_IF

(* 段 2：轴向速率、每转弧长与合成进给 *)
_fRpS := REAL_TO_LREAL(fSpindleRpm);
_fVzMmMin := fPitchMmRev * _fRpS;                        // mm/rev × r/min = mm/min
_fArcPerRev := 2.0 * DL_HEL_PI * fRadiusMm;              // 每转弧长 / Arc length per revolution
_fSumSq := fFeedProgMmMin * fFeedProgMmMin + _fVzMmMin * _fVzMmMin;
IF ((_fVzMmMin - _fVzMmMin) <> (_fVzMmMin - _fVzMmMin)) OR (_fSumSq < 0.0) THEN
    RETURN;                                              // 轴向速率 ±Inf 或平方和异常 / Non-finite axial rate
END_IF
fZPerRev := LREAL_TO_REAL(fPitchMmRev);
fHelixFeedMmMin := LREAL_TO_REAL(SQRT(_fSumSq));

(* 段 3：升角校验（螺距 > 每转弧长 ⇔ 升角 > 45°） *)
_uCode := 0;
IF fPitchMmRev > _fArcPerRev THEN _uCode := 5; END_IF

(* 段 4：结果复检 + 单一出口裁决（N4） *)
IF (fZPerRev <> fZPerRev) OR (fHelixFeedMmMin <> fHelixFeedMmMin)
   OR ((fHelixFeedMmMin - fHelixFeedMmMin) <> (fHelixFeedMmMin - fHelixFeedMmMin)) THEN
    fZPerRev := 0.0;  fHelixFeedMmMin := 0.0;  _uCode := 4;
END_IF
uErrId := _uCode;
IF _uCode = 0 THEN FC_DL_HelicalTurnAdvanceCalc := TRUE; END_IF
END_FUNCTION

(* ---- FC_DL_HoistSyncSpeedCalc.st ---- *)
(*
 * FC_DL_HoistSyncSpeedCalc | C2 | DL_Motion
 * 功能：双卷筒起升主从同步速度微调量与同步到位判定       单位：速度 [m/s]、增益 [1]、偏差 [m/s]
 * 工况边界：仅适用于主从同轴刚性/柔性双卷筒同步（不含位置闭环校正）；rTrimMaxMps 与 rDevLimitMps 须 >0 且有限，否则 xValid=FALSE 且微调量取 0；NaN/±Inf 一律拒算
 * 代数值回代：vMaster=0.50、vSlave=0.46、Kp=0.8、TrimMax=0.05、DevLimit=0.02 → dev=0.04、trim=0.032（未打限幅）、xInSync=FALSE（与 spec 回代行一致）
 * 开源溯源：clean-room 自研，未复制任何第三方代码（无外部来源）
 *)
FUNCTION FC_DL_HoistSyncSpeedCalc : BOOL
VAR_INPUT
    rVMasterMps  : REAL;             // 主卷筒速度给定 | master drum speed reference [m/s]
    rVSlaveMps   : REAL;             // 从卷筒速度反馈 | slave drum speed feedback [m/s]
    rKp          : REAL := 0.8;      // 偏差比例增益（无量纲）| proportional gain on the deviation [1]
    rTrimMaxMps  : REAL := 0.05;     // 从卷筒微调量限幅 | slave trim magnitude limit [m/s]
    rDevLimitMps : REAL := 0.02;     // 同步判定偏差阈 | in-sync deviation threshold [m/s]
END_VAR
VAR_OUTPUT
    rSlaveTrimMps  : REAL;           // 从卷筒速度微调量（已限幅）| slave speed trim after limiting [m/s]
    rDevMps        : REAL;           // 主从速度偏差（主−从）| master minus slave deviation [m/s]
    rAbsDevMps     : REAL;           // 偏差绝对值（判据与告警同源）| absolute deviation shared by the criterion and the alarm [m/s]
    xInSync        : BOOL;           // 同步到位 | in-sync flag
    xTrimSaturated : BOOL;           // 微调量已打限幅（信息级）| trim saturated, informational only
    xValid         : BOOL;           // 输出有效 | outputs valid
END_VAR
VAR
    xFinM   : BOOL;                  // 主速度有限性 | master speed is finite
    xFinS   : BOOL;                  // 从速度有限性 | slave speed is finite
    xFinKp  : BOOL;                  // 增益有限性 | gain is finite
    xFinMax : BOOL;                  // 限幅有限性 | trim limit is finite
    xFinDev : BOOL;                  // 判定阈有限性 | deviation threshold is finite
    rTrimRaw: REAL;                  // 未限幅微调量 | raw trim before limiting [m/s]
END_VAR

// 段1｜非有限闸（R19：非有限一律出口取 0 并置 xValid=FALSE）
xFinM := (rVMasterMps = rVMasterMps) AND ((rVMasterMps - rVMasterMps) = 0.0);
xFinS := (rVSlaveMps = rVSlaveMps) AND ((rVSlaveMps - rVSlaveMps) = 0.0);
xFinKp := (rKp = rKp) AND ((rKp - rKp) = 0.0);
xFinMax := (rTrimMaxMps = rTrimMaxMps) AND ((rTrimMaxMps - rTrimMaxMps) = 0.0);
xFinDev := (rDevLimitMps = rDevLimitMps) AND ((rDevLimitMps - rDevLimitMps) = 0.0);
IF (NOT xFinM) OR (NOT xFinS) OR (NOT xFinKp) OR (NOT xFinMax) OR (NOT xFinDev) THEN
    rSlaveTrimMps := 0.0;            // 安全值：不加微调，从卷筒按原给定 | safe value, no trim applied
    rDevMps := 0.0;
    rAbsDevMps := 0.0;
    xInSync := FALSE;                // 不可判定即判不同步，禁止联动起升 | not judgeable means out of sync
    xTrimSaturated := FALSE;
    xValid := FALSE;
    FC_DL_HoistSyncSpeedCalc := FALSE;
    RETURN;
END_IF

// 段2｜域闸：限幅与判定阈必须为正（LIMIT 边界必须有界）
IF (rTrimMaxMps <= 0.0) OR (rDevLimitMps <= 0.0) THEN
    rSlaveTrimMps := 0.0;
    rDevMps := 0.0;
    rAbsDevMps := 0.0;
    xInSync := FALSE;
    xTrimSaturated := FALSE;
    xValid := FALSE;
    FC_DL_HoistSyncSpeedCalc := FALSE;
    RETURN;
END_IF

// 段3｜算法：dev = 主 − 从；trim = LIMIT(−max, Kp*dev, max)；同步判据用未钳位的原始偏差
rDevMps := rVMasterMps - rVSlaveMps;
rAbsDevMps := ABS(rDevMps);                                // 判据与告警同源（R24）| criterion and alarm share the same source
rTrimRaw := rKp * rDevMps;
rSlaveTrimMps := LIMIT(-rTrimMaxMps, rTrimRaw, rTrimMaxMps);
xTrimSaturated := ABS(rTrimRaw) > rTrimMaxMps;             // 打限幅即置信息位 | flag saturation as information
xInSync := rAbsDevMps <= rDevLimitMps;                     // 用原始偏差判定，不受限幅影响 | judged on the raw deviation

// 段4｜出口
xValid := TRUE;
FC_DL_HoistSyncSpeedCalc := TRUE;
END_FUNCTION

(* ---- FC_DL_LaneDiverterAngleCalc.st ---- *)
(*
  ============================================================
  组件名 : FC_DL_LaneDiverterAngleCalc
  分类   : DL_Motion
  功能   : 道岔转角计算，由包件宽度与道间距求最小偏转角并折算通过时间与速度许可
  复杂度 : C2
  版本   : 1.0.0
  作者   : 道莅工业代码库工厂 / R81
  日期   : 2026-11-24
  开源溯源 : clean-room（no upstream）—— 依据公开工程公式自研，未复制任何上游实现
  红线自检 : R1 无GVL/R2 无物理地址/R3 纯IEC/R4 防除零/R5 双语注释
  接口说明 :
      最小转角 = ATAN(包件宽度 / 道间距)，ATAN 以弧度返回，再除以 0.0174533 折算为度。
      通过时间 = (包件长度/1000) / (线速度/60)，即长度折米后除以速度折 m/s。
      线速度不超过 60 m/min 判速度许可；速度为 0 时通过时间无定义，判无效。
  ============================================================
*)
FUNCTION FC_DL_LaneDiverterAngleCalc : BOOL
VAR_INPUT
    bEnable    : BOOL; // 使能：TRUE 时计算 / Enable: TRUE to compute
    bErr       : BOOL; // 外部故障：TRUE 时立即退出并置结果无效 / External fault: TRUE aborts with invalid result
    rPkgW_mm   : REAL; // 包件宽度，垂直于输送方向 [mm] / package width perpendicular to the conveying direction [millimetre]
    rPkgL_mm   : REAL; // 包件长度，沿输送方向 [mm] / package length along the conveying direction [millimetre]
    rLaneGap_mm : REAL; // 相邻道中心间距 [mm] / centre distance between adjacent lanes [millimetre]
    rSpeedMpm  : REAL; // 输送线速度 [m/min] / conveyor line speed [metre per minute]
END_VAR
VAR_OUTPUT
    rAngleRad : REAL; // 最小偏转角 [rad] / minimum divert angle [radian]
    rAngleDeg : REAL; // 最小偏转角 [度] / minimum divert angle [degree]
    rCrossTime_s : REAL; // 包件通过道岔所需时间 [s] / time for the package to cross the diverter [second]
    bSpeedOk  : BOOL; // 速度许可：TRUE 表示线速度不超过 60 m/min / speed permitted, TRUE when the line speed is within 60 metres per minute
    bValid    : BOOL; // 输出有效：TRUE 表示结果可用 / Output valid
END_VAR
VAR CONSTANT
    DL_R_MAX     : REAL := 3.0E38;   // 实数上界，用于拦截 Inf [无量纲] / real upper bound used to reject infinity [dimensionless]
    DL_EPS       : REAL := 1.0E-12;  // 除零判定阈值 [无量纲] / division guard threshold [dimensionless]
    DL_RAD_TO_DEG : REAL := 0.0174533; // 弧度转度系数 [度/rad] / radian to degree factor [degree per radian]
    DL_MM_TO_M   : REAL := 1000.0;   // 毫米折米系数 [mm/m] / millimetre to metre factor [millimetre per metre]
    DL_MIN_PER_S : REAL := 60.0;     // 每分钟秒数 [s/min] / seconds per minute [second per minute]
    DL_SPEED_OK  : REAL := 60.0;     // 允许的最高线速度 [m/min] / permitted maximum line speed [metre per minute]
    DL_SPEED_MAX : REAL := 600.0;    // 线速度合理上限 [m/min] / sanity upper bound of the line speed [metre per minute]
    DL_GAP_MIN   : REAL := 1.0;      // 道间距合理下限 [mm] / sanity lower bound of the lane gap [millimetre]
    DL_GAP_MAX   : REAL := 10000.0;  // 道间距合理上限 [mm] / sanity upper bound of the lane gap [millimetre]
    DL_SIZE_MAX  : REAL := 5000.0;   // 包件尺寸合理上限 [mm] / sanity upper bound of the package dimension [millimetre]
END_VAR
VAR
    _bFin    : BOOL := FALSE; // 输入有限性判定结果 / input finiteness verdict
    _rLenM   : REAL := 0.0;   // 包件长度折算米 [m] / package length in metre [metre]
    _rSpdMs  : REAL := 0.0;   // 线速度折算米每秒 [m/s] / line speed in metre per second [metre per second]
END_VAR

    // 段 1｜出口预置
    rAngleRad := 0.0;
    rAngleDeg := 0.0;
    rCrossTime_s := 0.0;
    bSpeedOk := FALSE;
    bValid := FALSE;
    // 段 2｜使能闸与外部故障闸
    IF NOT bEnable THEN
        RETURN;
    END_IF;
    IF bErr THEN
        RETURN;
    END_IF;
    // 段 3｜非有限闸
    _bFin := (rPkgW_mm = rPkgW_mm) AND (ABS(rPkgW_mm) <= DL_R_MAX) AND (rPkgL_mm = rPkgL_mm) AND (ABS(rPkgL_mm) <= DL_R_MAX) AND (rLaneGap_mm = rLaneGap_mm) AND (ABS(rLaneGap_mm) <= DL_R_MAX) AND (rSpeedMpm = rSpeedMpm) AND (ABS(rSpeedMpm) <= DL_R_MAX);
    IF NOT _bFin THEN
        RETURN;
    END_IF;
    // 段 4｜域闸：包件尺寸非负且合理，道间距在合理区间，速度严格为正且合理
    IF (rPkgW_mm < 0.0) OR (rPkgW_mm > DL_SIZE_MAX) OR (rPkgL_mm < 0.0) OR (rPkgL_mm > DL_SIZE_MAX) THEN
        RETURN;
    END_IF;
    IF (rLaneGap_mm < DL_GAP_MIN) OR (rLaneGap_mm > DL_GAP_MAX) THEN
        RETURN;
    END_IF;
    IF (ABS(rSpeedMpm) <= DL_EPS) OR (rSpeedMpm < 0.0) OR (rSpeedMpm > DL_SPEED_MAX) THEN
        RETURN;
    END_IF;
    // 段 5｜最小转角
    rAngleRad := ATAN(rPkgW_mm / rLaneGap_mm);
    rAngleDeg := rAngleRad / DL_RAD_TO_DEG;
    // 段 6｜通过时间：长度折米、速度折米每秒
    _rLenM := rPkgL_mm / DL_MM_TO_M;
    _rSpdMs := rSpeedMpm / DL_MIN_PER_S;
    IF ABS(_rSpdMs) <= DL_EPS THEN
        RETURN;
    END_IF;
    rCrossTime_s := _rLenM / _rSpdMs;
    // 段 7｜速度许可
    IF rSpeedMpm <= DL_SPEED_OK THEN
        bSpeedOk := TRUE;
    ELSE
        bSpeedOk := FALSE;
    END_IF;
    bValid := TRUE;
    FC_DL_LaneDiverterAngleCalc := bValid;
END_FUNCTION

(* ---- FC_DL_LineSpeedMatchRatio.st ---- *)
(*
  ============================================================
  组件名 : FC_DL_LineSpeedMatchRatio
  分类   : DL_Motion
  功能   : 主从线速匹配校验，由主从线速求实际速比并与设定速比比较给出偏差与匹配位
  复杂度 : C1
  版本   : 1.0.0
  作者   : 道莅工业代码库工厂 / R81
  日期   : 2026-11-24
  开源溯源 : clean-room（no upstream）—— 依据公开工程公式自研，未复制任何上游实现
  红线自检 : R1 无GVL/R2 无物理地址/R3 纯IEC/R4 防除零/R5 双语注释
  接口说明 :
      实际速比 = 从线速度 / 主线速度；偏差 = (实际速比 - 设定速比) / 设定速比 * 100。
      偏差绝对值不超过 2% 判匹配；主线静止时速比无定义，直接判无效而不是输出零速比。
  ============================================================
*)
FUNCTION FC_DL_LineSpeedMatchRatio : BOOL
VAR_INPUT
    bEnable    : BOOL; // 使能：TRUE 时校验 / Enable: TRUE to check
    bErr       : BOOL; // 外部故障：TRUE 时立即退出并置结果无效 / External fault: TRUE aborts with invalid result
    rMasterMpm : REAL; // 主线线速度 [m/min] / master line speed [metre per minute]
    rSlaveMpm  : REAL; // 从线线速度 [m/min] / slave line speed [metre per minute]
    rRatioSet  : REAL; // 设定速比，从线相对主线 [无量纲] / set speed ratio of slave over master [dimensionless]
END_VAR
VAR_OUTPUT
    rRatioAct : REAL; // 实际速比 [无量纲] / actual speed ratio [dimensionless]
    rDevPct   : REAL; // 速比相对偏差 [%] / relative speed ratio deviation [percent]
    bMatch    : BOOL; // 匹配：TRUE 表示偏差绝对值不超过 2% / matched, TRUE when the absolute deviation is within 2 percent
    bValid    : BOOL; // 输出有效：TRUE 表示结果可用 / Output valid
END_VAR
VAR CONSTANT
    DL_R_MAX   : REAL := 3.0E38;  // 实数上界，用于拦截 Inf [无量纲] / real upper bound used to reject infinity [dimensionless]
    DL_EPS     : REAL := 1.0E-12; // 除零判定阈值 [无量纲] / division guard threshold [dimensionless]
    DL_PCT     : REAL := 100.0;   // 百分数换算系数 [无量纲] / percentage scaling factor [dimensionless]
    DL_TOL_PCT : REAL := 2.0;     // 速比匹配允许偏差 [%] / permitted ratio deviation for a match [percent]
    DL_RATIO_MAX : REAL := 100.0; // 速比合理上限 [无量纲] / sanity upper bound of the speed ratio [dimensionless]
    DL_SPEED_MAX : REAL := 10000.0; // 线速度合理上限 [m/min] / sanity upper bound of the line speed [metre per minute]
END_VAR
VAR
    _bFin   : BOOL := FALSE; // 输入有限性判定结果 / input finiteness verdict
    _rAbsDev : REAL := 0.0;  // 偏差绝对值 [%] / absolute deviation [percent]
END_VAR

    // 段 1｜出口预置
    rRatioAct := 0.0;
    rDevPct := 0.0;
    bMatch := FALSE;
    bValid := FALSE;
    // 段 2｜使能闸与外部故障闸
    IF NOT bEnable THEN
        RETURN;
    END_IF;
    IF bErr THEN
        RETURN;
    END_IF;
    // 段 3｜非有限闸
    _bFin := (rMasterMpm = rMasterMpm) AND (ABS(rMasterMpm) <= DL_R_MAX) AND (rSlaveMpm = rSlaveMpm) AND (ABS(rSlaveMpm) <= DL_R_MAX) AND (rRatioSet = rRatioSet) AND (ABS(rRatioSet) <= DL_R_MAX);
    IF NOT _bFin THEN
        RETURN;
    END_IF;
    // 段 4｜域闸：主线速度严格为正，从线速度非负，设定速比严格为正
    IF (ABS(rMasterMpm) <= DL_EPS) OR (rMasterMpm < 0.0) OR (rMasterMpm > DL_SPEED_MAX) THEN
        RETURN;
    END_IF;
    IF (rSlaveMpm < 0.0) OR (rSlaveMpm > DL_SPEED_MAX) THEN
        RETURN;
    END_IF;
    IF (ABS(rRatioSet) <= DL_EPS) OR (rRatioSet < 0.0) OR (rRatioSet > DL_RATIO_MAX) THEN
        RETURN;
    END_IF;
    // 段 5｜实际速比
    rRatioAct := rSlaveMpm / rMasterMpm;
    // 段 6｜相对偏差
    rDevPct := (rRatioAct - rRatioSet) / rRatioSet * DL_PCT;
    // 段 7｜匹配判定
    _rAbsDev := ABS(rDevPct);
    IF _rAbsDev <= DL_TOL_PCT THEN
        bMatch := TRUE;
    ELSE
        bMatch := FALSE;
    END_IF;
    bValid := TRUE;
    FC_DL_LineSpeedMatchRatio := bValid;
END_FUNCTION

(* ---- FC_DL_MecanumWheelForwardCalc.st ---- *)
// FC_DL_MecanumWheelForwardCalc v1.0.0
// 开源溯源：clean-room 自研（族 DL_Motion，ST 生态实测 0 命中，无外部代码引入）
(*
  功能: 麦克纳姆轮正运动学 k = a + b：vx = (vFL+vFR+vRL+vRR)/4，
        vy = (−vFL+vFR+vRL−vRR)/4，ω = (−vFL+vFR−vRL+vRR)/(4k)；k 为唯一分母。
  邻件/码位: 与 FC_DL_MecanumWheelInverseCalc 构成正/逆一对（轮→底盘侧，供轮速实测校核）；
             16#0002_9202 = 域外或非有限拒收。
*)
FUNCTION FC_DL_MecanumWheelForwardCalc : REAL
VAR_INPUT
    fVelFL   : REAL := 0.0;     // 左前轮线速度 [m/s] / Front-left speed [m/s]
    fVelFR   : REAL := 0.0;     // 右前轮线速度 [m/s] / Front-right speed [m/s]
    fVelRL   : REAL := 0.0;     // 左后轮线速度 [m/s] / Rear-left speed [m/s]
    fVelRR   : REAL := 0.0;     // 右后轮线速度 [m/s] / Rear-right speed [m/s]
    fHalfLen : REAL := 0.3;     // 半轴距 a [m]，纵向半跨 / Half wheelbase [m]
    fHalfWid : REAL := 0.25;    // 半轮距 b [m]，横向半跨 / Half track [m]
END_VAR
VAR_OUTPUT
    fVx      : REAL;            // 车体纵向速度 [m/s]，前正 / Longitudinal velocity [m/s]
    fVy      : REAL;            // 车体横向速度 [m/s]，左正 / Lateral velocity [m/s]
    fOmega   : REAL;            // 车体自转角速度 [rad/s] / Body yaw rate [rad/s]
    bValid   : BOOL;            // 结果有效回执 [-] / Result validity receipt
    uErrorId : UDINT;           // 事件码，0 = 无事件 / Event code
END_VAR
VAR
    fK : REAL := 0.0;           // 合成力臂 k = a + b [m] / Combined lever arm [m]
END_VAR
// 段 0：全路径出口安全缺省（三出口一律缺省）/ Safe defaults on all outlets
fVx := 0.0;                     // 纵向速度缺省零 / Longitudinal default zero
fVy := 0.0;                     // 横向速度缺省零 / Lateral default zero
fOmega := 0.0;                  // 角速度缺省零 / Yaw rate default zero
bValid := FALSE;                // 有效回执预清 / Validity preset clear
uErrorId := 16#0000;            // 事件码预清 / Event code preset clear
FC_DL_MecanumWheelForwardCalc := 0.0;   // 返回值缺省零（镜像纵向速度）/ Return default zero
// 段 1：非有限闸（四轮速 + 两几何量全枚举）/ Non-finite gate over all inputs
IF (fVelFL <> fVelFL) OR (fVelFR <> fVelFR) OR (fVelRL <> fVelRL) OR (fVelRR <> fVelRR)
   OR (fHalfLen <> fHalfLen) OR (fHalfWid <> fHalfWid)
   OR (ABS(fVelFL) >= 3.0E38) OR (ABS(fVelFR) >= 3.0E38) OR (ABS(fVelRL) >= 3.0E38)
   OR (ABS(fVelRR) >= 3.0E38) OR (ABS(fHalfLen) >= 3.0E38) OR (ABS(fHalfWid) >= 3.0E38) THEN
    uErrorId := 16#0002_9202;   // 入参非有限拒收 / Non-finite input reject
    RETURN;
END_IF
// 段 2：域闸（k 为正，ω 分母非零）/ Domain gate, R4 divide-by-zero guard
fK := fHalfLen + fHalfWid;      // 合成力臂 / Combined lever arm
IF fK <= 1.0E-6 THEN
    uErrorId := 16#0002_9202;   // 力臂非正，转向不可解 / Non-positive arm, yaw unsolvable
    RETURN;
END_IF
// 段 3：主计算（四轮线性组合）/ Main computation
fVx := (fVelFL + fVelFR + fVelRL + fVelRR) / 4.0;                   // 纵向速度均值 / Longitudinal mean
fVy := (-fVelFL + fVelFR + fVelRL - fVelRR) / 4.0;                  // 横向带符号组合 / Lateral signed sum
fOmega := (-fVelFL + fVelFR - fVelRL + fVelRR) / (4.0 * fK);        // 角速度除以力臂 / Yaw over arm
// 段 4：出口闸（三输出各做非有限复核）/ Outlet gate
IF (fVx <> fVx) OR (fVy <> fVy) OR (fOmega <> fOmega)
   OR (ABS(fVx) >= 3.0E38) OR (ABS(fVy) >= 3.0E38) OR (ABS(fOmega) >= 3.0E38) THEN
    fVx := 0.0;                 // 复核失败回缺省 / Fallback on recheck failure
    fVy := 0.0;                 // 复核失败回缺省 / Fallback on recheck failure
    fOmega := 0.0;              // 复核失败回缺省 / Fallback on recheck failure
    uErrorId := 16#0002_9202;   // 出口非有限拒收 / Output non-finite reject
    RETURN;
END_IF
bValid := TRUE;                 // 有效回执 / Validity receipt
FC_DL_MecanumWheelForwardCalc := fVx;   // 返回值镜像纵向速度 / Return mirrors longitudinal speed
END_FUNCTION

(* ---- FC_DL_MecanumWheelInverseCalc.st ---- *)
// FC_DL_MecanumWheelInverseCalc v1.0.0
// 开源溯源：clean-room 自研（族 DL_Motion，ST 生态实测 0 命中，无外部代码引入）
(*
  功能: 麦克纳姆轮逆运动学 k = a + b：vFL = vx − vy − ωk，vFR = vx + vy + ωk，
        vRL = vx + vy − ωk，vRR = vx − vy + ωk；fOmegaTotal 为四轮回算角速度自检。
  邻件/码位: 与 FC_DL_MecanumWheelForwardCalc 构成逆/正一对；16#0002_9201 = 域外或非有限拒收。
*)
FUNCTION FC_DL_MecanumWheelInverseCalc : REAL
VAR_INPUT
    fVx      : REAL := 0.0;     // 车体纵向速度 vx [m/s]，前正 / Longitudinal velocity [m/s]
    fVy      : REAL := 0.0;     // 车体横向速度 vy [m/s]，左正 / Lateral velocity [m/s]
    fOmega   : REAL := 0.0;     // 自转角速度 ω [rad/s]，逆时针正 / Yaw rate [rad/s]
    fRadius  : REAL := 0.05;    // 轮半径 [m]，域 >= 1e-3 / Wheel radius [m]
    fHalfLen : REAL := 0.3;     // 半轴距 a [m]，纵向半跨 / Half wheelbase [m]
    fHalfWid : REAL := 0.25;    // 半轮距 b [m]，横向半跨 / Half track [m]
END_VAR
VAR_OUTPUT
    fVelFL      : REAL;         // 左前轮线速度 [m/s] / Front-left speed [m/s]
    fVelFR      : REAL;         // 右前轮线速度 [m/s] / Front-right speed [m/s]
    fVelRL      : REAL;         // 左后轮线速度 [m/s] / Rear-left speed [m/s]
    fVelRR      : REAL;         // 右后轮线速度 [m/s] / Rear-right speed [m/s]
    fOmegaTotal : REAL;         // 四轮回算角速度 [rad/s] / Recomposed yaw rate [rad/s]
    bOverSpeed  : BOOL;         // 超速告警，仅告警不否决 [-] / Over-speed warning only
    bValid      : BOOL;         // 结果有效回执 [-] / Result validity receipt
    uErrorId    : UDINT;        // 事件码，0 = 无事件 / Event code
END_VAR
VAR
    fK : REAL := 0.0;           // 合成力臂 k = a + b [m] / Combined lever arm [m]
END_VAR
// 段 0：全路径出口安全缺省（不回灌入参）/ Safe defaults, inputs never echoed back
fVelFL := 0.0;                  // 左前轮速缺省零 / Front-left default zero
fVelFR := 0.0;                  // 右前轮速缺省零 / Front-right default zero
fVelRL := 0.0;                  // 左后轮速缺省零 / Rear-left default zero
fVelRR := 0.0;                  // 右后轮速缺省零 / Rear-right default zero
fOmegaTotal := 0.0;             // 回算角速度缺省零 / Recomposed yaw default zero
bOverSpeed := FALSE;            // 超速告警预清 / Over-speed preset clear
bValid := FALSE;                // 有效回执预清 / Validity preset clear
uErrorId := 16#0000;            // 事件码预清 / Event code preset clear
FC_DL_MecanumWheelInverseCalc := 0.0;   // 返回值缺省零（镜像左前轮速）/ Return default zero
// 段 1：非有限闸（六入参全枚举）/ Non-finite gate over all six inputs
IF (fVx <> fVx) OR (fVy <> fVy) OR (fOmega <> fOmega) OR (fRadius <> fRadius)
   OR (fHalfLen <> fHalfLen) OR (fHalfWid <> fHalfWid)
   OR (ABS(fVx) >= 3.0E38) OR (ABS(fVy) >= 3.0E38) OR (ABS(fOmega) >= 3.0E38)
   OR (ABS(fRadius) >= 3.0E38) OR (ABS(fHalfLen) >= 3.0E38) OR (ABS(fHalfWid) >= 3.0E38) THEN
    uErrorId := 16#0002_9201;   // 入参非有限拒收 / Non-finite input reject
    RETURN;
END_IF
// 段 2：域闸（半径下界 + 力臂为正，防除零）/ Domain gate, R4 divide-by-zero guard
fK := fHalfLen + fHalfWid;      // 合成力臂 / Combined lever arm
IF (fRadius < 1.0E-3) OR (fK <= 1.0E-6) THEN
    uErrorId := 16#0002_9201;   // 半径近零或力臂非正（几何不可解）/ Domain violation
    RETURN;
END_IF
// 段 3：主计算（四轮逆解，ωk 为旋转切向分量）/ Main computation
fVelFL := fVx - fVy - fOmega * fK;                                  // 左前轮 / Front-left wheel
fVelFR := fVx + fVy + fOmega * fK;                                  // 右前轮 / Front-right wheel
fVelRL := fVx + fVy - fOmega * fK;                                  // 左后轮 / Rear-left wheel
fVelRR := fVx - fVy + fOmega * fK;                                  // 右后轮 / Rear-right wheel
fOmegaTotal := (fVelFR + fVelRL - fVelFL - fVelRR) / (4.0 * fK);    // 四轮回算角速度自检 / Recomposed yaw
// 段 4：出口闸（非有限复核 + 超速告警）/ Outlet gate
IF (fVelFL <> fVelFL) OR (fVelFR <> fVelFR) OR (fVelRL <> fVelRL) OR (fVelRR <> fVelRR)
   OR (fOmegaTotal <> fOmegaTotal) OR (ABS(fOmegaTotal) >= 3.0E38) THEN
    fVelFL := 0.0;              // 复核失败回缺省 / Fallback on recheck failure
    fVelFR := 0.0;              // 复核失败回缺省 / Fallback on recheck failure
    fVelRL := 0.0;              // 复核失败回缺省 / Fallback on recheck failure
    fVelRR := 0.0;              // 复核失败回缺省 / Fallback on recheck failure
    fOmegaTotal := 0.0;         // 复核失败回缺省 / Fallback on recheck failure
    uErrorId := 16#0002_9201;   // 出口非有限拒收 / Output non-finite reject
    RETURN;
END_IF
IF (ABS(fVelFL) > 3.0) OR (ABS(fVelFR) > 3.0) OR (ABS(fVelRL) > 3.0) OR (ABS(fVelRR) > 3.0) THEN
    bOverSpeed := TRUE;         // 超速告警，仅标记不否决 / Over-speed warning, no veto
END_IF
bValid := TRUE;                 // 有效回执 / Validity receipt
FC_DL_MecanumWheelInverseCalc := fVelFL;    // 返回值镜像左前轮速 / Return mirrors front-left
END_FUNCTION

(* ---- FC_DL_PurePursuitCurvatureCalc.st ---- *)
// FC_DL_PurePursuitCurvatureCalc v1.0.0
// 开源溯源：clean-room 自研（族 DL_Motion，ST 生态实测 0 命中，无外部代码引入）
(*
  功能: 纯跟踪曲率律 Ld = MAX(fLookAhead, fMinLook)，alpha = ATAN2(y, x) 以
        ATAN(y/x) + 四象限修正实现（规避方言 ATAN2），κ = 2·SIN(alpha)/Ld。
  邻件/码位: 与 FC_DL_StanleySteerAngleCalc 同为跟踪律（预瞄点几何 vs 偏差反馈）；
             16#0002_9204 = 非有限、预瞄近零或目标点重合拒收。
*)
FUNCTION FC_DL_PurePursuitCurvatureCalc : REAL
VAR_INPUT
    fTargetX   : REAL := 1.0;       // 预瞄点车体坐标 X [m]，前正 / Look-ahead X [m]
    fTargetY   : REAL := 0.0;       // 预瞄点车体坐标 Y [m]，左正 / Look-ahead Y [m]
    fLookAhead : REAL := 1.0;       // 预瞄距离 [m]，域 > 0 / Look-ahead distance [m]
    fMinLook   : REAL := 0.3;       // 最小预瞄距离 [m] / Minimum look-ahead [m]
END_VAR
VAR_OUTPUT
    fCurvature : REAL;              // 期望曲率 κ [1/m]，左转为正 / Desired curvature [1/m]
    fAlpha     : REAL;              // 预瞄角 alpha [rad]，左转为正 / Look-ahead angle [rad]
    bValid     : BOOL;              // 结果有效回执 [-] / Result validity receipt
    uErrorId   : UDINT;             // 事件码，0 = 无事件 / Event code
END_VAR
VAR
    fPi     : REAL := 3.14159265358979; // 圆周率常量 [rad] / Pi constant [rad]
    fHalfPi : REAL := 1.5707963267949;  // 半圆周率 [rad] / Half pi constant [rad]
    fLd     : REAL := 0.0;              // 生效预瞄距离 [m] / Effective look-ahead [m]
END_VAR
// 段 0：全路径出口安全缺省（曲率零 = 直行）/ Safe defaults, zero curvature means straight
fCurvature := 0.0;              // 曲率缺省零 / Curvature default zero
fAlpha := 0.0;                  // 预瞄角缺省零 / Alpha default zero
bValid := FALSE;                // 有效回执预清 / Validity preset clear
uErrorId := 16#0000;            // 事件码预清 / Event code preset clear
FC_DL_PurePursuitCurvatureCalc := 0.0;  // 返回值缺省零 / Return default zero
// 段 1：非有限闸（四入参全枚举）/ Non-finite gate over all inputs
IF (fTargetX <> fTargetX) OR (fTargetY <> fTargetY)
   OR (fLookAhead <> fLookAhead) OR (fMinLook <> fMinLook)
   OR (ABS(fTargetX) >= 3.0E38) OR (ABS(fTargetY) >= 3.0E38)
   OR (ABS(fLookAhead) >= 3.0E38) OR (ABS(fMinLook) >= 3.0E38) THEN
    uErrorId := 16#0002_9204;   // 入参非有限拒收 / Non-finite input reject
    RETURN;
END_IF
// 段 2：域闸（预瞄取大后仍须为正 + 目标点不与原点重合）/ Domain gate
fLd := fLookAhead;                                              // 先取预瞄距离 / Take look-ahead first
IF fMinLook > fLd THEN
    fLd := fMinLook;                                            // 提升到最小预瞄 / Raise to minimum
END_IF
IF (fLd <= 1.0E-3) OR ((ABS(fTargetX) + ABS(fTargetY)) < 1.0E-6) THEN
    uErrorId := 16#0002_9204;   // 预瞄近零或目标点重合原点 / Degenerate look-ahead or target
    RETURN;
END_IF
// 段 3：主计算（ATAN + 四象限修正替代 ATAN2）/ Main computation
IF ABS(fTargetX) < 1.0E-9 THEN                                  // X 近零需定纵轴 / Axis branch
    IF fTargetY >= 0.0 THEN
        fAlpha := fHalfPi;                                      // 正纵轴 / Positive vertical axis
    ELSE
        fAlpha := -fHalfPi;                                     // 负纵轴 / Negative vertical axis
    END_IF
ELSE
    fAlpha := ATAN(fTargetY / fTargetX);                        // 主值分支 / Principal branch
    IF fTargetX < 0.0 THEN                                      // 左半平面补 π / Left half-plane fix
        IF fTargetY >= 0.0 THEN
            fAlpha := fAlpha + fPi;                             // 第二象限 / Second quadrant
        ELSE
            fAlpha := fAlpha - fPi;                             // 第三象限 / Third quadrant
        END_IF
    END_IF
END_IF
fCurvature := 2.0 * SIN(fAlpha) / fLd;                          // κ = 2·sin(alpha)/Ld / Curvature law
// 段 4：出口闸（双输出非有限复核）/ Outlet gate
IF (fCurvature <> fCurvature) OR (fAlpha <> fAlpha)
   OR (ABS(fCurvature) >= 3.0E38) OR (ABS(fAlpha) >= 3.0E38) THEN
    fCurvature := 0.0;          // 复核失败回缺省 / Fallback on recheck failure
    fAlpha := 0.0;              // 复核失败回缺省 / Fallback on recheck failure
    uErrorId := 16#0002_9204;   // 出口非有限拒收 / Output non-finite reject
    RETURN;
END_IF
bValid := TRUE;                 // 有效回执 / Validity receipt
FC_DL_PurePursuitCurvatureCalc := fCurvature;   // 返回值镜像曲率 / Return mirrors curvature
END_FUNCTION

(* ---- FC_DL_ResolverAmpImbalance.st ---- *)
(* ===========================================================================
   组件名   : FC_DL_ResolverAmpImbalance
   分类     : DL_Motion / 旋转变压器幅值不平衡
   一句话   : 计算 sin/cos 两路幅值不平衡度百分比并判定是否超限
   复杂度   : 1        版本 : v1.0.0        日期 : 2026-11-24
   开源溯源 : 无（clean-room 自研，未借鉴任何开源实现）
   输入契约 : fSinAmp 正弦路峰值幅值 [V]；fCosAmp 余弦路峰值幅值 [V]
              fLimitPct 不平衡度限值 [%]
   输出契约 : 返回值 = 不平衡度 [%]（|A−B| / 均值 × 100）
              xOverLimit 是否超限；xValid 输入有效；fMeanAmp 两路均值 [V]
   修改记录 : v1.0.0 2026-11-24 初版
   =========================================================================== *)

FUNCTION FC_DL_ResolverAmpImbalance : REAL
VAR_INPUT
    fSinAmp : REAL;                    // 正弦路峰值幅值 [V] | sine channel amplitude [V]
    fCosAmp : REAL;                    // 余弦路峰值幅值 [V] | cosine channel amplitude [V]
    fLimitPct : REAL := 5.0;           // 不平衡度限值 [%] | imbalance limit [%]
END_VAR
VAR_OUTPUT
    xOverLimit : BOOL;                 // 不平衡超限标志 | imbalance over limit
    xValid : BOOL;                     // 输入有效标志 | inputs valid flag
    fMeanAmp : REAL;                   // 两路均值幅值 [V] | mean amplitude [V]
END_VAR
VAR
    _fSum : REAL;                      // 两路幅值之和 [V] | sum of amplitudes [V]
    _fDiff : REAL;                      // 两路幅值之差 [V] | difference of amplitudes [V]
    _fPct : REAL;                      // 不平衡度 [%] | imbalance [%]
END_VAR

// ---- 输出预置：防止调用方读到未初始化值 ----
xOverLimit := FALSE;
xValid := FALSE;
fMeanAmp := 0.0;
_fPct := 0.0;
FC_DL_ResolverAmpImbalance := 0.0;

// ---- 非有限值拦截 ----
IF (fSinAmp <> fSinAmp) OR ((fSinAmp - fSinAmp) <> (fSinAmp - fSinAmp)) THEN
    RETURN;
END_IF
IF (fCosAmp <> fCosAmp) OR ((fCosAmp - fCosAmp) <> (fCosAmp - fCosAmp)) THEN
    RETURN;
END_IF
IF (fLimitPct <> fLimitPct) OR ((fLimitPct - fLimitPct) <> (fLimitPct - fLimitPct)) THEN
    RETURN;
END_IF

_fSum := ABS(fSinAmp) + ABS(fCosAmp);
fMeanAmp := _fSum * 0.5;

// ---- 零幅值保护：均值为零时不平衡度无定义，判无效 ----
IF fMeanAmp > 0.000000001 THEN
    _fDiff := ABS(ABS(fSinAmp) - ABS(fCosAmp));
    _fPct := _fDiff / fMeanAmp * 100.0;            // 分母已守卫
    xValid := TRUE;
    IF fLimitPct > 0.0 THEN
        xOverLimit := (_fPct > fLimitPct);         // 用大于比较，不做浮点等值判定
    END_IF
END_IF

FC_DL_ResolverAmpImbalance := _fPct;
END_FUNCTION

(* ---- FC_DL_ResolverAngleDecode.st ---- *)
(* ===========================================================================
   组件名   : FC_DL_ResolverAngleDecode
   分类     : DL_Motion / 旋转变压器角度解算
   一句话   : 由 sin/cos 两路幅值解算机械角，arctan2 采用分段线性近似加象限修正
   复杂度   : 2        版本 : v1.0.0        日期 : 2026-11-24
   开源溯源 : 无（clean-room 自研，未借鉴任何开源实现）
   输入契约 : fSin 正弦路瞬时值 [V]；fCos 余弦路瞬时值 [V]；fAmpMin 最小有效合成幅值 [V]
   输出契约 : 返回值 = 机械角 [rad]，范围 [0, 2π)；xValid 解算有效
              fAmplitude 合成幅值 [V]；fRatioNorm 归一化插值量 0..1（诊断用）
   算法说明 : atan(t) ≈ t / (1 + 0.28086·t^2)，t 为小值/大值（0..1），误差优于 0.005 rad
              象限修正按 atan2 恒等式：|x|≥|y| 取 base，否则取 π/2−base；x<0 取 π−θ，y<0 取 −θ
   修改记录 : v1.0.0 2026-11-24 初版
   =========================================================================== *)

FUNCTION FC_DL_ResolverAngleDecode : REAL
VAR_INPUT
    fSin : REAL;                       // 正弦路瞬时值 [V] | sine channel value [V]
    fCos : REAL;                       // 余弦路瞬时值 [V] | cosine channel value [V]
    fAmpMin : REAL := 0.1;             // 最小有效合成幅值 [V] | min valid amplitude [V]
END_VAR
VAR_OUTPUT
    xValid : BOOL;                     // 解算有效标志 | decode valid flag
    fAmplitude : REAL;                 // 合成幅值 [V] | resultant amplitude [V]
    fRatioNorm : REAL;                 // 归一化插值量 0..1 | normalized ratio 0..1
END_VAR
VAR
    _fAbsSin : REAL;                   // 正弦绝对值 [V] | absolute sine [V]
    _fAbsCos : REAL;                   // 余弦绝对值 [V] | absolute cosine [V]
    _fMin : REAL;                      // 两路绝对值较小者 [V] | smaller magnitude [V]
    _fMax : REAL;                      // 两路绝对值较大者 [V] | larger magnitude [V]
    _fT : REAL;                        // 小/大 归一化比 0..1 | small/large ratio 0..1
    _fBase : REAL;                     // 基准角 [rad] | base angle [rad]
    _fOut : REAL;                      // 结果角 [rad] | result angle [rad]
END_VAR

// ---- 输出预置：任何提前返回路径都不会留下未初始化值 ----
xValid := FALSE;
fAmplitude := 0.0;
fRatioNorm := 0.0;
FC_DL_ResolverAngleDecode := 0.0;

// ---- 非有限值拦截：NaN 用自反比较，Inf 用 (x-x)<>(x-x) ----
IF ((fSin <> fSin) OR ((fSin - fSin) <> (fSin - fSin))) THEN
    RETURN;
END_IF
IF ((fCos <> fCos) OR ((fCos - fCos) <> (fCos - fCos))) THEN
    RETURN;
END_IF

_fAbsSin := ABS(fSin);
_fAbsCos := ABS(fCos);
fAmplitude := SQRT(fSin * fSin + fCos * fCos);

// ---- 幅值为零保护：合成幅值不足则角度不可信 ----
IF (fAmpMin <= 0.0) OR (fAmplitude < fAmpMin) THEN
    RETURN;
END_IF
xValid := TRUE;

// ---- 归一化：小值 / 大值 落在 0..1，分母由幅值门限保证非零 ----
_fMax := MAX(_fAbsSin, _fAbsCos);
_fMin := MIN(_fAbsSin, _fAbsCos);
IF _fMax < 0.000000001 THEN
    xValid := FALSE;                                // 双路同时近零，再兜底一次
    RETURN;
END_IF
_fT := _fMin / _fMax;                               // 分母已守卫
fRatioNorm := _fT;

// ---- atan 分段线性近似（t 在 0..1，结果在 0..π/4） ----
_fBase := _fT / (1.0 + 0.28086 * _fT * _fT);

// ---- 象限修正：先按 |x| 与 |y| 的大小关系选基准轴 ----
IF _fAbsCos >= _fAbsSin THEN
    _fOut := _fBase;                                // 以余弦轴为基准
ELSE
    _fOut := 1.570796327 - _fBase;                  // π/2 − base
END_IF

// ---- 符号修正：x<0 折到第二/三象限，y<0 取负角 ----
IF fCos < 0.0 THEN
    _fOut := 3.141592654 - _fOut;
END_IF
IF fSin < 0.0 THEN
    _fOut := -_fOut;
END_IF

// ---- 归一化到 [0, 2π) ----
IF _fOut < 0.0 THEN
    _fOut := _fOut + 6.283185307;
END_IF
IF _fOut >= 6.283185307 THEN
    _fOut := _fOut - 6.283185307;
END_IF

FC_DL_ResolverAngleDecode := _fOut;
END_FUNCTION

(* ---- FC_DL_ResolverElecAngleUnwrap.st ---- *)
(* ===========================================================================
   组件名   : FC_DL_ResolverElecAngleUnwrap
   分类     : DL_Motion / 旋转变压器电角度解卷绕
   一句话   : 跨 0/2π 边界时累加圈数，输出连续电角度与圈数
   复杂度   : 2        版本 : v1.0.0        日期 : 2026-11-24
   开源溯源 : 无（clean-room 自研，未借鉴任何开源实现）
   输入契约 : fAngleNow 本拍电角度 [rad] 0..2π；fAnglePrev 上拍电角度 [rad] 0..2π
              iTurnPrev 上拍累计圈数
   输出契约 : 返回值 = 连续电角度 [rad]（可超出 0..2π）
              iTurns 本拍累计圈数；fDelta 解卷绕后电角增量 [rad]；xValid 输入有效
   修改记录 : v1.0.0 2026-11-24 初版
   =========================================================================== *)

FUNCTION FC_DL_ResolverElecAngleUnwrap : REAL
VAR_INPUT
    fAngleNow : REAL;                  // 本拍电角度 [rad] | current electrical angle [rad]
    fAnglePrev : REAL;                 // 上拍电角度 [rad] | previous electrical angle [rad]
    iTurnPrev : INT := 0;              // 上拍累计圈数 | previous turn count
END_VAR
VAR_OUTPUT
    iTurns : INT;                      // 本拍累计圈数 | current turn count
    fDelta : REAL;                     // 解卷绕后增量 [rad] | unwrapped delta [rad]
    xValid : BOOL;                     // 输入有效标志 | inputs valid flag
END_VAR
VAR
    _fD : REAL;                        // 本拍角差 [rad] | angle difference [rad]
    _iT : INT;                         // 累计圈数工作值 | turn count working value
END_VAR

// ---- 输出预置 ----
iTurns := 0;
fDelta := 0.0;
xValid := FALSE;
FC_DL_ResolverElecAngleUnwrap := 0.0;

// ---- 非有限值拦截 ----
IF (fAngleNow <> fAngleNow) OR ((fAngleNow - fAngleNow) <> (fAngleNow - fAngleNow)) THEN
    RETURN;
END_IF
IF (fAnglePrev <> fAnglePrev) OR ((fAnglePrev - fAnglePrev) <> (fAnglePrev - fAnglePrev)) THEN
    RETURN;
END_IF

// ---- 圈数钳位：防止长时间运行后整型溢出 ----
_iT := iTurnPrev;
IF _iT > 1000000 THEN
    _iT := 1000000;
ELSIF _iT < -1000000 THEN
    _iT := -1000000;
END_IF

// ---- 解卷绕：正向跨零（差 < −π）圈数 +1，反向跨零（差 > π）圈数 −1 ----
_fD := fAngleNow - fAnglePrev;
IF _fD > 3.141592654 THEN
    _fD := _fD - 6.283185307;                      // 反向跨零补偿
    _iT := _iT - 1;
ELSIF _fD < -3.141592654 THEN
    _fD := _fD + 6.283185307;                      // 正向跨零补偿
    _iT := _iT + 1;
END_IF

// ---- 圈数二次钳位：补偿后仍须落在可表范围内 ----
IF _iT > 1000000 THEN
    _iT := 1000000;
ELSIF _iT < -1000000 THEN
    _iT := -1000000;
END_IF

fDelta := _fD;
iTurns := _iT;
xValid := TRUE;

// ---- 连续角 = 圈数 × 2π + 本拍角 ----
FC_DL_ResolverElecAngleUnwrap := INT_TO_REAL(_iT) * 6.283185307 + fAngleNow;
END_FUNCTION

(* ---- FC_DL_ResolverExcitationPhaseChk.st ---- *)
(* ===========================================================================
   组件名   : FC_DL_ResolverExcitationPhaseChk
   分类     : DL_Motion / 旋转变压器励磁相位校验
   一句话   : 校验励磁与输出的相位差是否命中期望值，并据此判定接线相序是否反接
   复杂度   : 2        版本 : v1.0.0        日期 : 2026-11-24
   开源溯源 : 无（clean-room 自研，未借鉴任何开源实现）
   输入契约 : fExcPhase 励磁相位 [rad]；fOutPhase 输出相位 [rad]
              fExpectedDiff 期望相位差 [rad]；fTol 容差 [rad]
   输出契约 : 返回值 = 卷绕到 (−π, π] 的实测相位差 [rad]
              xPhaseOk 相位差落在期望值容差内；xSeqReversed 判为相序反接（差 180°）
              xValid 输入有效
   修改记录 : v1.0.0 2026-11-24 初版
   =========================================================================== *)

FUNCTION FC_DL_ResolverExcitationPhaseChk : REAL
VAR_INPUT
    fExcPhase : REAL;                  // 励磁相位 [rad] | excitation phase [rad]
    fOutPhase : REAL;                  // 输出相位 [rad] | output phase [rad]
    fExpectedDiff : REAL := 0.0;       // 期望相位差 [rad] | expected phase difference [rad]
    fTol : REAL := 0.2;                // 相位容差 [rad] | phase tolerance [rad]
END_VAR
VAR_OUTPUT
    xPhaseOk : BOOL;                   // 相位差合格 | phase difference acceptable
    xSeqReversed : BOOL;               // 相序反接（差 180°） | wiring reversed (180 deg)
    xValid : BOOL;                     // 输入有效标志 | inputs valid flag
END_VAR
VAR
    _fDiff : REAL;                     // 卷绕后相位差 [rad] | wrapped phase difference [rad]
    _fErrFwd : REAL;                   // 与期望值的偏差（正接） [rad] | error, forward wiring [rad]
    _fErrRev : REAL;                   // 与期望值的偏差（反接） [rad] | error, reversed wiring [rad]
    _fTmp : REAL;                      // 卷绕中间量 [rad] | wrap intermediate [rad]
END_VAR

// ---- 输出预置 ----
xPhaseOk := FALSE;
xSeqReversed := FALSE;
xValid := FALSE;
FC_DL_ResolverExcitationPhaseChk := 0.0;

// ---- 非有限值拦截 ----
IF (fExcPhase <> fExcPhase) OR ((fExcPhase - fExcPhase) <> (fExcPhase - fExcPhase)) THEN
    RETURN;
END_IF
IF (fOutPhase <> fOutPhase) OR ((fOutPhase - fOutPhase) <> (fOutPhase - fOutPhase)) THEN
    RETURN;
END_IF
IF (fTol <> fTol) OR ((fTol - fTol) <> (fTol - fTol)) OR (fTol <= 0.0) THEN
    RETURN;
END_IF

// ---- 实测相位差并卷绕到 (−π, π] ----
_fDiff := fOutPhase - fExcPhase;
IF _fDiff > 1000000.0 THEN
    _fDiff := 1000000.0;                           // 上限钳位，防 TRUNC 溢出
ELSIF _fDiff < -1000000.0 THEN
    _fDiff := -1000000.0;
END_IF
_fDiff := _fDiff - 6.283185307 * TRUNC(_fDiff / 6.283185307);
IF _fDiff > 3.141592654 THEN
    _fDiff := _fDiff - 6.283185307;
ELSIF _fDiff <= -3.141592654 THEN
    _fDiff := _fDiff + 6.283185307;
END_IF
FC_DL_ResolverExcitationPhaseChk := _fDiff;

// ---- 正接偏差：实测差 − 期望差，再卷绕 ----
_fTmp := _fDiff - fExpectedDiff;
IF _fTmp > 3.141592654 THEN
    _fTmp := _fTmp - 6.283185307;
ELSIF _fTmp <= -3.141592654 THEN
    _fTmp := _fTmp + 6.283185307;
END_IF
_fErrFwd := ABS(_fTmp);                            // 绝对值即偏差幅度

// ---- 反接偏差：正接偏差再叠加 180° ----
_fTmp := _fTmp + 3.141592654;
IF _fTmp > 3.141592654 THEN
    _fTmp := _fTmp - 6.283185307;
ELSIF _fTmp <= -3.141592654 THEN
    _fTmp := _fTmp + 6.283185307;
END_IF
_fErrRev := ABS(_fTmp);

// ---- 判定：容差比较一律用小于等于，不做浮点等值判定 ----
IF _fErrFwd <= fTol THEN
    xPhaseOk := TRUE;                              // 正接合格
ELSIF _fErrRev <= fTol THEN
    xSeqReversed := TRUE;                          // 差 180° 判为相序反接
END_IF
xValid := TRUE;
END_FUNCTION

(* ---- FC_DL_ResolverOffsetTrim.st ---- *)
(* ===========================================================================
   组件名   : FC_DL_ResolverOffsetTrim
   分类     : DL_Motion / 旋转变压器零位标定
   一句话   : 记录安装零位偏置并按偏置修正输出角，两模式共用同一取模归一逻辑
   复杂度   : 1        版本 : v1.0.0        日期 : 2026-11-24
   开源溯源 : 无（clean-room 自研，未借鉴任何开源实现）
   输入契约 : fAngleRaw 原始机械角 [rad]；fOffset 已存偏置 [rad]；fAngleRef 参考零位 [rad]
              xCapture TRUE=标定本拍（记录偏置），FALSE=应用偏置
   输出契约 : 返回值 = 修正后机械角 [rad]，范围 [0, 2π)；fOffsetOut 生效偏置 [rad]
              xValid 输入有效
   修改记录 : v1.0.0 2026-11-24 初版
   =========================================================================== *)

FUNCTION FC_DL_ResolverOffsetTrim : REAL
VAR_INPUT
    fAngleRaw : REAL;                  // 原始机械角 [rad] | raw mechanical angle [rad]
    fOffset : REAL;                    // 已存零位偏置 [rad] | stored zero offset [rad]
    fAngleRef : REAL := 0.0;           // 参考零位 [rad] | reference zero angle [rad]
    xCapture : BOOL;                   // TRUE=标定模式 | TRUE=capture mode
END_VAR
VAR_OUTPUT
    fOffsetOut : REAL;                 // 生效偏置 [rad] | effective offset [rad]
    xValid : BOOL;                     // 输入有效标志 | inputs valid flag
END_VAR
VAR
    _fTmp : REAL;                      // 取模中间量 [rad] | modulo intermediate [rad]
    _fCyc : REAL;                      // 圈数整数值 | integer turns value
    _fOut : REAL;                      // 修正角 [rad] | corrected angle [rad]
END_VAR

// ---- 输出预置 ----
fOffsetOut := 0.0;
xValid := FALSE;
FC_DL_ResolverOffsetTrim := 0.0;

// ---- 非有限值拦截 ----
IF (fAngleRaw <> fAngleRaw) OR ((fAngleRaw - fAngleRaw) <> (fAngleRaw - fAngleRaw)) THEN
    RETURN;
END_IF
IF (fOffset <> fOffset) OR ((fOffset - fOffset) <> (fOffset - fOffset)) THEN
    RETURN;
END_IF
IF (fAngleRef <> fAngleRef) OR ((fAngleRef - fAngleRef) <> (fAngleRef - fAngleRef)) THEN
    RETURN;
END_IF

IF xCapture THEN
    // ---- 标定模式：偏置 = 原始角 − 参考零位，取模到 [0, 2π) ----
    _fTmp := fAngleRaw - fAngleRef;
    IF _fTmp > 1000000.0 THEN
        _fTmp := 1000000.0;                        // 上限钳位，防 TRUNC 溢出
    ELSIF _fTmp < -1000000.0 THEN
        _fTmp := -1000000.0;
    END_IF
    _fCyc := TRUNC(_fTmp / 6.283185307);           // 常量分母，非零
    _fTmp := _fTmp - 6.283185307 * _fCyc;
    IF _fTmp < 0.0 THEN
        _fTmp := _fTmp + 6.283185307;
    END_IF
    IF _fTmp >= 6.283185307 THEN
        _fTmp := _fTmp - 6.283185307;
    END_IF
    fOffsetOut := _fTmp;
    _fOut := fAngleRaw;                            // 标定拍不改变已解算角
    xValid := TRUE;
ELSE
    // ---- 应用模式：偏置取模后从原始角扣除 ----
    _fTmp := fOffset;
    IF _fTmp > 1000000.0 THEN
        _fTmp := 1000000.0;
    ELSIF _fTmp < -1000000.0 THEN
        _fTmp := -1000000.0;
    END_IF
    _fCyc := TRUNC(_fTmp / 6.283185307);
    _fTmp := _fTmp - 6.283185307 * _fCyc;
    IF _fTmp < 0.0 THEN
        _fTmp := _fTmp + 6.283185307;
    END_IF
    IF _fTmp >= 6.283185307 THEN
        _fTmp := _fTmp - 6.283185307;
    END_IF
    fOffsetOut := _fTmp;

    _fOut := fAngleRaw - _fTmp;
    IF _fOut < 0.0 THEN
        _fOut := _fOut + 6.283185307;              // 负角归一
    END_IF
    IF _fOut >= 6.283185307 THEN
        _fOut := _fOut - 6.283185307;
    END_IF
    xValid := TRUE;
END_IF

FC_DL_ResolverOffsetTrim := _fOut;
END_FUNCTION

(* ---- FC_DL_ResolverPolePairAngle.st ---- *)
(* ===========================================================================
   组件名   : FC_DL_ResolverPolePairAngle
   分类     : DL_Motion / 旋转变压器电角度换算
   一句话   : 由机械角与极对数换算电角度，含取模与负角归一化处理
   复杂度   : 2        版本 : v1.0.0        日期 : 2026-11-24
   开源溯源 : 无（clean-room 自研，未借鉴任何开源实现）
   输入契约 : fMechAngle 机械角 [rad]；iPolePairs 极对数 1..64；fMechOffset 机械零位偏置 [rad]
   输出契约 : 返回值 = 电角度 [rad]，范围 [0, 2π)；fElecTurns 电角累计整圈数
              xValid 输入有效
   修改记录 : v1.0.0 2026-11-24 初版
   =========================================================================== *)

FUNCTION FC_DL_ResolverPolePairAngle : REAL
VAR_INPUT
    fMechAngle : REAL;                 // 机械角 [rad] | mechanical angle [rad]
    iPolePairs : INT := 1;             // 极对数 1..64 | pole pairs 1..64
    fMechOffset : REAL := 0.0;         // 机械零位偏置 [rad] | mechanical zero offset [rad]
END_VAR
VAR_OUTPUT
    fElecTurns : REAL;                 // 电角整圈数（截断值） | electrical whole turns
    xValid : BOOL;                     // 输入有效标志 | inputs valid flag
END_VAR
VAR
    _fRaw : REAL;                      // 未归一电角度 [rad] | unnormalized electrical angle [rad]
    _fCyc : REAL;                      // 整圈数值 | whole turns value
    _fOut : REAL;                      // 归一化电角度 [rad] | normalized electrical angle [rad]
    _iPP : INT;                        // 钳位后极对数 | clamped pole pairs
END_VAR

// ---- 输出预置 ----
fElecTurns := 0.0;
xValid := FALSE;
FC_DL_ResolverPolePairAngle := 0.0;

// ---- 非有限值拦截 ----
IF (fMechAngle <> fMechAngle) OR ((fMechAngle - fMechAngle) <> (fMechAngle - fMechAngle)) THEN
    RETURN;
END_IF
IF (fMechOffset <> fMechOffset) OR ((fMechOffset - fMechOffset) <> (fMechOffset - fMechOffset)) THEN
    RETURN;
END_IF

// ---- 极对数钳位：上限 64 防乘后数值过大，下限 1 防退化为零角 ----
_iPP := iPolePairs;
IF _iPP < 1 THEN
    _iPP := 1;
ELSIF _iPP > 64 THEN
    _iPP := 64;
END_IF

// ---- 电角度 = （机械角 − 零位偏置）× 极对数 ----
_fRaw := (fMechAngle - fMechOffset) * INT_TO_REAL(_iPP);
IF _fRaw > 1000000.0 THEN
    _fRaw := 1000000.0;                            // 上限钳位，防 TRUNC 溢出
ELSIF _fRaw < -1000000.0 THEN
    _fRaw := -1000000.0;
END_IF

// ---- 取模归一：先截断圈数再扣余量，避免正向循环累减 ----
_fCyc := TRUNC(_fRaw / 6.283185307);               // 常量分母，非零
_fOut := _fRaw - 6.283185307 * _fCyc;              // 余量落在 (−2π, 2π)

// ---- 负角归一化到 [0, 2π) ----
IF _fOut < 0.0 THEN
    _fOut := _fOut + 6.283185307;
END_IF
IF _fOut >= 6.283185307 THEN
    _fOut := _fOut - 6.283185307;                  // 浮点余量兜底，单次修正足够
END_IF

fElecTurns := _fCyc;
xValid := TRUE;
FC_DL_ResolverPolePairAngle := _fOut;
END_FUNCTION

(* ---- FC_DL_ResolverSpeedCalc.st ---- *)
(* ===========================================================================
   组件名   : FC_DL_ResolverSpeedCalc
   分类     : DL_Motion / 旋转变压器测速
   一句话   : 由相邻两拍角度差分解算转速，含跨零解卷绕与一阶低通滤波（状态由调用方持有）
   复杂度   : 2        版本 : v1.0.0        日期 : 2026-11-24
   开源溯源 : 无（clean-room 自研，未借鉴任何开源实现）
   输入契约 : fAngleNow 本拍角度 [rad] 0..2π；fAnglePrev 上拍角度 [rad] 0..2π
              fDtSec 采样周期 [s]；fSpeedPrev 上拍滤波后转速 [rad/s]；fLpfAlpha 低通系数 0..1
   输出契约 : 返回值 = 本拍滤波后转速 [rad/s]；fDeltaUnwrapped 解卷绕后角增量 [rad]
              xWrapFlag 本拍发生跨零解卷绕；xValid 输入有效
   修改记录 : v1.0.0 2026-11-24 初版
   =========================================================================== *)

FUNCTION FC_DL_ResolverSpeedCalc : REAL
VAR_INPUT
    fAngleNow : REAL;                  // 本拍角度 [rad] 0..2π | current angle [rad]
    fAnglePrev : REAL;                 // 上拍角度 [rad] 0..2π | previous angle [rad]
    fDtSec : REAL := 0.004;            // 采样周期 [s] | sample period [s]
    fSpeedPrev : REAL;                 // 上拍滤波后转速 [rad/s] | previous filtered speed [rad/s]
    fLpfAlpha : REAL := 0.2;           // 一阶低通系数 0..1 | first order lpf alpha
END_VAR
VAR_OUTPUT
    fDeltaUnwrapped : REAL;            // 解卷绕后角增量 [rad] | unwrapped angle delta [rad]
    fSpeedRaw : REAL;                  // 原始转速 [rad/s] | raw speed [rad/s]
    xWrapFlag : BOOL;                  // 是否发生跨零解卷绕 | wrap corrected flag
    xValid : BOOL;                     // 输入有效标志 | inputs valid flag
END_VAR
VAR
    _fDelta : REAL;                    // 角增量 [rad] | angle delta [rad]
    _fDt : REAL;                       // 钳位后采样周期 [s] | clamped dt [s]
    _fAlpha : REAL;                    // 钳位后低通系数 | clamped alpha
    _fSpeed : REAL;                    // 滤波后转速 [rad/s] | filtered speed [rad/s]
END_VAR

// ---- 输出预置 ----
fDeltaUnwrapped := 0.0;
fSpeedRaw := 0.0;
xWrapFlag := FALSE;
xValid := FALSE;
FC_DL_ResolverSpeedCalc := 0.0;

// ---- 非有限值拦截 ----
IF (fAngleNow <> fAngleNow) OR ((fAngleNow - fAngleNow) <> (fAngleNow - fAngleNow)) THEN
    RETURN;
END_IF
IF (fAnglePrev <> fAnglePrev) OR ((fAnglePrev - fAnglePrev) <> (fAnglePrev - fAnglePrev)) THEN
    RETURN;
END_IF
IF (fSpeedPrev <> fSpeedPrev) OR ((fSpeedPrev - fSpeedPrev) <> (fSpeedPrev - fSpeedPrev)) THEN
    RETURN;
END_IF

// ---- 周期钳位：防止零除与超大解算步长 ----
_fDt := fDtSec;
IF _fDt < 0.000001 THEN
    _fDt := 0.000001;
ELSIF _fDt > 0.2 THEN
    _fDt := 0.2;
END_IF

// ---- 角度跨零解卷绕：增量超出 ±π 即判为绕圈并补偿 2π ----
_fDelta := fAngleNow - fAnglePrev;
IF _fDelta > 3.141592654 THEN
    _fDelta := _fDelta - 6.283185307;              // 正向跨零
    xWrapFlag := TRUE;
ELSIF _fDelta < -3.141592654 THEN
    _fDelta := _fDelta + 6.283185307;              // 反向跨零
    xWrapFlag := TRUE;
END_IF
fDeltaUnwrapped := _fDelta;

// ---- 原始转速：分母已守卫 ----
fSpeedRaw := _fDelta / _fDt;

// ---- 一阶低通：系数钳位到 0..1 ----
_fAlpha := fLpfAlpha;
IF _fAlpha < 0.0 THEN
    _fAlpha := 0.0;
ELSIF _fAlpha > 1.0 THEN
    _fAlpha := 1.0;
END_IF
_fSpeed := fSpeedPrev + _fAlpha * (fSpeedRaw - fSpeedPrev);

xValid := TRUE;
FC_DL_ResolverSpeedCalc := _fSpeed;
END_FUNCTION

(* ---- FC_DL_RollerSlipRatioCalc.st ---- *)
(*
  ============================================================
  组件名 : FC_DL_RollerSlipRatioCalc
  分类   : DL_Motion
  功能   : 辊筒打滑率计算，由输送带速与辊面线速求相对打滑比例并给出打滑报警
  复杂度 : C1
  版本   : 1.0.0
  作者   : 道莅工业代码库工厂 / R81
  日期   : 2026-11-24
  开源溯源 : clean-room（no upstream）—— 依据公开工程公式自研，未复制任何上游实现
  红线自检 : R1 无GVL/R2 无物理地址/R3 纯IEC/R4 防除零/R5 双语注释
  接口说明 :
      打滑率 = (辊面线速 - 带速) / 辊面线速 * 100，限幅 -100~100。
      正值表示带速低于辊面速度即打滑，负值表示带速快于辊面速度即被拖动。
      打滑率绝对值超过 5% 置打滑报警；辊面线速为零时打滑率无定义，判无效。
  ============================================================
*)
FUNCTION FC_DL_RollerSlipRatioCalc : BOOL
VAR_INPUT
    bEnable    : BOOL; // 使能：TRUE 时计算 / Enable: TRUE to compute
    bErr       : BOOL; // 外部故障：TRUE 时立即退出并置结果无效 / External fault: TRUE aborts with invalid result
    rBeltMpm   : REAL; // 输送带实际线速度 [m/min] / actual belt speed [metre per minute]
    rRollerMpm : REAL; // 辊筒表面线速度 [m/min] / roller surface speed [metre per minute]
END_VAR
VAR_OUTPUT
    rSlipPct   : REAL; // 打滑率，限幅 -100~100 [%] / slip ratio clamped between minus 100 and 100 [percent]
    bSlipAlarm : BOOL; // 打滑报警：TRUE 表示打滑率绝对值超过 5% / slip alarm, TRUE when the absolute slip ratio exceeds 5 percent
    bValid     : BOOL; // 输出有效：TRUE 表示结果可用 / Output valid
END_VAR
VAR CONSTANT
    DL_R_MAX    : REAL := 3.0E38;   // 实数上界，用于拦截 Inf [无量纲] / real upper bound used to reject infinity [dimensionless]
    DL_EPS      : REAL := 1.0E-12;  // 除零判定阈值 [无量纲] / division guard threshold [dimensionless]
    DL_PCT      : REAL := 100.0;    // 百分数换算系数 [无量纲] / percentage scaling factor [dimensionless]
    DL_SLIP_HI  : REAL := 100.0;    // 打滑率限幅上限 [%] / upper clamp of the slip ratio [percent]
    DL_SLIP_LO  : REAL := -100.0;   // 打滑率限幅下限 [%] / lower clamp of the slip ratio [percent]
    DL_ALARM_PCT : REAL := 5.0;     // 打滑报警门限 [%] / slip alarm threshold [percent]
    DL_SPEED_MAX : REAL := 10000.0; // 线速度合理上限 [m/min] / sanity upper bound of the line speed [metre per minute]
END_VAR
VAR
    _bFin   : BOOL := FALSE; // 输入有限性判定结果 / input finiteness verdict
    _rRaw   : REAL := 0.0;   // 限幅前打滑率 [%] / raw slip ratio before clamping [percent]
    _rAbs   : REAL := 0.0;   // 打滑率绝对值 [%] / absolute slip ratio [percent]
END_VAR

    // 段 1｜出口预置
    rSlipPct := 0.0;
    bSlipAlarm := FALSE;
    bValid := FALSE;
    // 段 2｜使能闸与外部故障闸
    IF NOT bEnable THEN
        RETURN;
    END_IF;
    IF bErr THEN
        RETURN;
    END_IF;
    // 段 3｜非有限闸
    _bFin := (rBeltMpm = rBeltMpm) AND (ABS(rBeltMpm) <= DL_R_MAX) AND (rRollerMpm = rRollerMpm) AND (ABS(rRollerMpm) <= DL_R_MAX);
    IF NOT _bFin THEN
        RETURN;
    END_IF;
    // 段 4｜域闸：辊面线速严格为正，带速非负，两者均不超过合理上限
    IF (ABS(rRollerMpm) <= DL_EPS) OR (rRollerMpm < 0.0) OR (rRollerMpm > DL_SPEED_MAX) THEN
        RETURN;
    END_IF;
    IF (rBeltMpm < 0.0) OR (rBeltMpm > DL_SPEED_MAX) THEN
        RETURN;
    END_IF;
    // 段 5｜打滑率原值
    _rRaw := (rRollerMpm - rBeltMpm) / rRollerMpm * DL_PCT;
    // 段 6｜限幅
    IF _rRaw < DL_SLIP_LO THEN
        rSlipPct := DL_SLIP_LO;
    ELSIF _rRaw > DL_SLIP_HI THEN
        rSlipPct := DL_SLIP_HI;
    ELSE
        rSlipPct := _rRaw;
    END_IF;
    // 段 7｜报警判定
    _rAbs := ABS(rSlipPct);
    IF _rAbs > DL_ALARM_PCT THEN
        bSlipAlarm := TRUE;
    ELSE
        bSlipAlarm := FALSE;
    END_IF;
    bValid := TRUE;
    FC_DL_RollerSlipRatioCalc := bValid;
END_FUNCTION

(* ---- FC_DL_RotFeedInvTimeCalc.st ---- *)
(* ============================================================
   DL_Motion / FC_DL_RotFeedInvTimeCalc ｜ v1.0.0 ｜ 2026-11-25
   功能：旋转轴进给率双向换算与限幅。正向 INV_TIME[1/min]×每转角度[deg/rev]
         = deg/min；反向按限幅比例折算等效每转进给 fFeedPerRev[deg/rev]
   边界：INV≤0 / 每转角度≤0 / 上限≤0 → 码 1/2/3；非有限 → 码 4；三者均写 0 出口（N1/N3）
   依赖：仅 IEC 61131-3（MIN） ｜ 溯源：DLF-A-RTCP（内部原创线）
   ============================================================ *)
FUNCTION FC_DL_RotFeedInvTimeCalc : BOOL
VAR_INPUT
    fInvTimeVal    : LREAL;  // INV_TIME 编程值，域 > 0 [1/min] / Inverse time value per minute
    fDegPerRev     : LREAL;  // 每转对应角度（分度轴 360）[deg/rev] / Degrees per revolution
    fFeedMaxDegMin : LREAL;  // 允许进给上限，域 > 0 [deg/min] / Allowed feed ceiling
END_VAR
VAR_OUTPUT
    fFeedDegMin : LREAL;  // 限幅后进给率 [deg/min] / Limited feed rate
    fFeedPerRev : LREAL;  // 折算后每转进给 [deg/rev] / Effective advance per revolution
    uErrId      : UDINT;  // 出口码 0/1/2/3/4 [-] / Outlet code
    bLimited    : BOOL;   // 本拍被上限钳制 [-] / Feed clamped by the ceiling
END_VAR
VAR
    _fRaw : LREAL;  // 未限幅进给率 = INV × 每转角度 [deg/min] / Unlimited feed rate
END_VAR
VAR CONSTANT
    DL_RFI_EPS : LREAL := 1.0E-9;  // 判零与判等容差 [deg/min] / Zero and equality tolerance
END_VAR

(* 段 0：出口预置安全侧（进给 0 即停转，N3） *)
FC_DL_RotFeedInvTimeCalc := FALSE;
fFeedDegMin := 0.0;  fFeedPerRev := 0.0;  bLimited := TRUE;  uErrId := 4;

(* 段 1：非有限闸 + 三域闸 *)
IF (fInvTimeVal <> fInvTimeVal) OR (fDegPerRev <> fDegPerRev) OR (fFeedMaxDegMin <> fFeedMaxDegMin) THEN
    RETURN;
END_IF
IF fInvTimeVal <= 0.0 THEN uErrId := 1; RETURN; END_IF
IF fDegPerRev <= 0.0 THEN uErrId := 2; RETURN; END_IF
IF fFeedMaxDegMin <= 0.0 THEN uErrId := 3; RETURN; END_IF

(* 段 2：正向换算 INV[1/min] × 每转角度[deg/rev] = [deg/min] *)
_fRaw := fInvTimeVal * fDegPerRev;
IF (_fRaw <> _fRaw) OR ((_fRaw - _fRaw) <> (_fRaw - _fRaw)) THEN RETURN; END_IF

(* 段 3：单侧限幅（进给恒非负），标志与出口同源 *)
IF _fRaw > fFeedMaxDegMin + DL_RFI_EPS THEN
    fFeedDegMin := fFeedMaxDegMin;  bLimited := TRUE;
ELSE
    fFeedDegMin := _fRaw;  bLimited := FALSE;
END_IF

(* 段 4：反向折算（除子 _fRaw 已证 > 0） + 单一出口裁决（N4） *)
fFeedPerRev := fDegPerRev * (fFeedDegMin / _fRaw);
IF (fFeedPerRev <> fFeedPerRev) OR ((fFeedPerRev - fFeedPerRev) <> (fFeedPerRev - fFeedPerRev)) THEN
    fFeedDegMin := 0.0;  fFeedPerRev := 0.0;  bLimited := TRUE;  uErrId := 4;  RETURN;
END_IF
uErrId := 0;  FC_DL_RotFeedInvTimeCalc := TRUE;
END_FUNCTION

(* ---- FC_DL_RtcpPivotOffsetCalc.st ---- *)
(* ============================================================
   DL_Motion / FC_DL_RtcpPivotOffsetCalc ｜ v1.0.0 ｜ 2026-11-25
   功能：RTCP 摆动轴枢轴偏置在工件坐标系的三向分量 [mm]；
         刀具轴单位向量 v=(sinB·cosA, −sinA, cosA·cosB)，偏移 = L·(v − (0,0,1))
   边界：摆角先折叠到 (−180°,180°]，超 8 次折叠即钳位并置 bFolded；
         枢轴长度≤0 或非有限 → 三分量同步写 0、返回 FALSE（N1）
   依赖：仅 IEC 61131-3（SIN / COS） ｜ 溯源：DLF-A-RTCP（内部原创线）
   ============================================================ *)
FUNCTION FC_DL_RtcpPivotOffsetCalc : BOOL
VAR_INPUT
    fPivotLenMm : LREAL;  // 枢轴长度（主轴端面到摆心）[mm] / Pivot length from face to swivel center
    fTiltADeg   : REAL;   // 摆动轴 A 角（绕 X）[deg] / Swivel axis A angle about X
    fTiltBDeg   : REAL;   // 摆动轴 B 角（绕 Y）[deg] / Swivel axis B angle about Y
END_VAR
VAR_OUTPUT
    fDxMm   : REAL;   // 枢轴偏置 X 分量 [mm] / Pivot offset in X
    fDyMm   : REAL;   // 枢轴偏置 Y 分量 [mm] / Pivot offset in Y
    fDzMm   : REAL;   // 枢轴偏置 Z 分量 [mm] / Pivot offset in Z
    bFolded : BOOL;   // 摆角发生 360° 折叠 [-] / Angle folding happened
END_VAR
VAR
    _fA   : LREAL;  // 折叠后 A 角 [deg] / Folded angle of axis A
    _fB   : LREAL;  // 折叠后 B 角 [deg] / Folded angle of axis B
    _fAr  : LREAL;  // A 角弧度值 [rad] / Angle A in radians
    _fBr  : LREAL;  // B 角弧度值 [rad] / Angle B in radians
    _nIdx : INT;    // 折叠循环索引（上限 8 防死循环）[-] / Bounded fold loop index
END_VAR
VAR CONSTANT
    DL_RTPV_PI : LREAL := 3.14159265358979324;  // 圆周率（LREAL 全精度）[-] / Pi at full precision
END_VAR

(* 段 0：出口预置安全侧 + 非有限闸 *)
FC_DL_RtcpPivotOffsetCalc := FALSE;
fDxMm := 0.0;  fDyMm := 0.0;  fDzMm := 0.0;  bFolded := FALSE;
IF (fPivotLenMm <> fPivotLenMm) OR (fTiltADeg <> fTiltADeg) OR (fTiltBDeg <> fTiltBDeg) THEN
    RETURN;
END_IF
IF (fPivotLenMm - fPivotLenMm) <> (fPivotLenMm - fPivotLenMm) THEN RETURN; END_IF
IF fPivotLenMm <= 0.0 THEN RETURN; END_IF               // 组态非法：三分量保持 0

(* 段 1：摆角折叠到 (−180°,180°]，次数有界（N2：折叠结果为当拍值） *)
_fA := REAL_TO_LREAL(fTiltADeg);
_fB := REAL_TO_LREAL(fTiltBDeg);
FOR _nIdx := 1 TO 8 DO
    IF _fA > 180.0 THEN
        _fA := _fA - 360.0;  bFolded := TRUE;
    ELSIF _fA <= -180.0 THEN
        _fA := _fA + 360.0;  bFolded := TRUE;
    END_IF
    IF _fB > 180.0 THEN
        _fB := _fB - 360.0;  bFolded := TRUE;
    ELSIF _fB <= -180.0 THEN
        _fB := _fB + 360.0;  bFolded := TRUE;
    END_IF
END_FOR
IF _fA > 180.0 THEN _fA := 180.0; END_IF                 // 超 8 次折叠仍越域：钳位
IF _fA < -180.0 THEN _fA := -180.0; END_IF
IF _fB > 180.0 THEN _fB := 180.0; END_IF
IF _fB < -180.0 THEN _fB := -180.0; END_IF

(* 段 2：角度换算弧度，三向分量 = L × (v − 单位 Z) *)
_fAr := _fA * DL_RTPV_PI / 180.0;
_fBr := _fB * DL_RTPV_PI / 180.0;
fDxMm := LREAL_TO_REAL(fPivotLenMm * (SIN(_fBr) * COS(_fAr)));
fDyMm := LREAL_TO_REAL(fPivotLenMm * (0.0 - SIN(_fAr)));
fDzMm := LREAL_TO_REAL(fPivotLenMm * (COS(_fAr) * COS(_fBr) - 1.0));

(* 段 3：结果复检 + 单一出口裁决（N4） *)
IF (fDxMm <> fDxMm) OR (fDyMm <> fDyMm) OR (fDzMm <> fDzMm) THEN
    fDxMm := 0.0;  fDyMm := 0.0;  fDzMm := 0.0;  RETURN;
END_IF
FC_DL_RtcpPivotOffsetCalc := TRUE;
END_FUNCTION

(* ---- FC_DL_RtcpTrackingErrCalc.st ---- *)
(* ============================================================
   DL_Motion / FC_DL_RtcpTrackingErrCalc ｜ v1.0.0 ｜ 2026-11-25
   功能：RTCP 下编程点与实绩点三维偏差模长 √(dX²+dY²+dZ²) [mm]：
         分量 = 编程 − 实绩；模长超 5 mm 门限置码 1（供上层降速/停机）
   边界：分量非有限 → 模长 0、码 2（N1：判据与出口同源改写）；门限≤0 → 码 3；
         平方和溢出为非有限 → 同走码 2
   依赖：仅 IEC 61131-3（SQRT） ｜ 溯源：DLF-A-RTCP（内部原创线）
   ============================================================ *)
FUNCTION FC_DL_RtcpTrackingErrCalc : BOOL
VAR_INPUT
    fProgXmm : LREAL;  // 编程点 X [mm] / Programmed point X
    fProgYmm : LREAL;  // 编程点 Y [mm] / Programmed point Y
    fProgZmm : LREAL;  // 编程点 Z [mm] / Programmed point Z
    fActXmm  : LREAL;  // 实绩点 X [mm] / Actual point X
    fActYmm  : LREAL;  // 实绩点 Y [mm] / Actual point Y
    fActZmm  : LREAL;  // 实绩点 Z [mm] / Actual point Z
END_VAR
VAR_OUTPUT
    fErrMagMm : LREAL;  // 三维偏差模长 [mm] / Magnitude of the deviation
    uErrId    : UDINT;  // 出口码 0 正常 / 1 超差 / 2 非有限 / 3 门限非法 [-] / Outlet code
END_VAR
VAR
    _fDx  : LREAL;  // X 向分量 [mm] / Deviation component in X
    _fDy  : LREAL;  // Y 向分量 [mm] / Deviation component in Y
    _fDz  : LREAL;  // Z 向分量 [mm] / Deviation component in Z
    _fSum : LREAL;  // 三分量平方和 [mm²] / Sum of squared components
END_VAR
VAR CONSTANT
    DL_RTE_LIMIT : LREAL := 5.0;  // 跟踪误差门限 [mm] / Tracking error threshold
END_VAR

(* 段 0：出口预置安全侧 *)
FC_DL_RtcpTrackingErrCalc := FALSE;
fErrMagMm := 0.0;  uErrId := 2;

(* 段 1：非有限闸（六个入参全量枚举） *)
IF (fProgXmm <> fProgXmm) OR (fProgYmm <> fProgYmm) OR (fProgZmm <> fProgZmm)
   OR (fActXmm <> fActXmm) OR (fActYmm <> fActYmm) OR (fActZmm <> fActZmm) THEN
    RETURN;
END_IF
IF ((fProgXmm - fProgXmm) <> (fProgXmm - fProgXmm)) THEN RETURN; END_IF

(* 段 2：三分量与模长 *)
_fDx := fProgXmm - fActXmm;  _fDy := fProgYmm - fActYmm;  _fDz := fProgZmm - fActZmm;
_fSum := _fDx * _fDx + _fDy * _fDy + _fDz * _fDz;
IF (_fSum <> _fSum) OR ((_fSum - _fSum) <> (_fSum - _fSum)) OR (_fSum < 0.0) THEN
    RETURN;                                              // 平方和非有限或为负：结构性兜底
END_IF
fErrMagMm := SQRT(_fSum);

(* 段 3：门限判据（门限先过域闸，禁先夹量程再判超限）与出口裁决（N4） *)
IF DL_RTE_LIMIT <= 0.0 THEN
    uErrId := 3;
ELSIF fErrMagMm > DL_RTE_LIMIT THEN
    uErrId := 1;                                         // 超差：模长照给，返回 FALSE
ELSE
    uErrId := 0;  FC_DL_RtcpTrackingErrCalc := TRUE;
END_IF
END_FUNCTION

(* ---- FC_DL_SagFeedLimitCalc.st ---- *)
(* ============================================================
   DL_Motion / FC_DL_SagFeedLimitCalc ｜ v1.0.0 ｜ 2026-11-25
   功能：按允许弦高、向心加速度上限与采样周期反解进给上限 [mm/min]：
         v_sag = √(8·R·e)/T，v_acc = √(a·R)，取小值 ×60
   边界：半径≤0 / 弦高≤0 / 加速度≤0 / 周期=0 或非有限 → 上限写 0、bLimited=TRUE（N1/N3）
         bLimited=TRUE 表示被弦高约束压死（向心约束更紧时为 FALSE）
   依赖：仅 IEC 61131-3（SQRT / MIN / TIME_TO_REAL） ｜ 溯源：DLF-A-RTCP（内部原创线）
   ============================================================ *)
FUNCTION FC_DL_SagFeedLimitCalc : BOOL
VAR_INPUT
    fSagTolMm   : LREAL;  // 允许弦高（垂度）容差，域 > 0 [mm] / Allowed chord sag tolerance
    fRadiusMm   : LREAL;  // 路径曲率半径，域 > 0 [mm] / Path curvature radius
    fAccMaxMmS2 : LREAL;  // 向心加速度上限，域 > 0 [mm/s²] / Centripetal acceleration ceiling
    tCycle      : TIME;   // 插补采样周期，域 > 0 [ms] / Interpolation sampling period
END_VAR
VAR_OUTPUT
    fFeedMaxMmMin : LREAL;  // 进给率上限 [mm/min] / Feed rate ceiling
    bLimited      : BOOL;   // 输出被弦高约束压死 [-] / Output bound by the sag constraint
END_VAR
VAR
    _fTSec : LREAL;  // 采样周期换算值 [s] / Sampling period in seconds
    _fVSag : LREAL;  // 弦高约束允许速度 [mm/s] / Speed allowed by the sag constraint
    _fVAcc : LREAL;  // 向心约束允许速度 [mm/s] / Speed allowed by the centripetal constraint
END_VAR
VAR CONSTANT
    DL_SAG_MS_PER_S : LREAL := 1000.0;  // 毫秒 → 秒换算系数 [ms/s] / Milliseconds per second
END_VAR

(* 段 0：出口预置安全侧（上限 0 = 禁止运动，N3） *)
FC_DL_SagFeedLimitCalc := FALSE;
fFeedMaxMmMin := 0.0;  bLimited := TRUE;

(* 段 1：非有限闸 + 四域闸 *)
IF (fSagTolMm <> fSagTolMm) OR (fRadiusMm <> fRadiusMm) OR (fAccMaxMmS2 <> fAccMaxMmS2) THEN
    RETURN;
END_IF
IF (fRadiusMm <= 0.0) OR (fSagTolMm <= 0.0) OR (fAccMaxMmS2 <= 0.0) THEN RETURN; END_IF
_fTSec := TIME_TO_REAL(tCycle) / DL_SAG_MS_PER_S;        // ms → s
IF _fTSec <= 0.0 THEN RETURN; END_IF

(* 段 2：两约束允许速度（开方前已证根号内 > 0） *)
_fVSag := SQRT(8.0 * fRadiusMm * fSagTolMm) / _fTSec;
_fVAcc := SQRT(fAccMaxMmS2 * fRadiusMm);

(* 段 3：取小值、判约束源，同步落进给上限（N4 单段裁决） *)
IF _fVSag < _fVAcc THEN
    fFeedMaxMmMin := _fVSag * 60.0;  bLimited := TRUE;   // 弦高约束更紧
ELSE
    fFeedMaxMmMin := _fVAcc * 60.0;  bLimited := FALSE;  // 向心约束更紧
END_IF

(* 段 4：结果复检（出口闸位于最后一次赋值之后） *)
IF (fFeedMaxMmMin <> fFeedMaxMmMin)
   OR ((fFeedMaxMmMin - fFeedMaxMmMin) <> (fFeedMaxMmMin - fFeedMaxMmMin)) THEN
    fFeedMaxMmMin := 0.0;  bLimited := TRUE;  RETURN;
END_IF
FC_DL_SagFeedLimitCalc := TRUE;
END_FUNCTION

(* ---- FC_DL_SkateWheelLoadCalc.st ---- *)
(*
  ============================================================
  组件名 : FC_DL_SkateWheelLoadCalc
  分类   : DL_Motion
  功能   : 滑板轮载荷分配计算，按重心纵向偏移求前后轴占比并折算前轴单轮载荷
  复杂度 : C2
  版本   : 1.0.0
  作者   : 道莅工业代码库工厂 / R81
  日期   : 2026-11-24
  开源溯源 : clean-room（no upstream）—— 依据公开工程公式自研，未复制任何上游实现
  红线自检 : R1 无GVL/R2 无物理地址/R3 纯IEC/R4 防除零/R5 双语注释
  接口说明 :
      前轴占比 = 0.5 + 重心偏移 / 轴距，限幅 0.1~0.9，防止极端重心把全部载荷压到单轴。
      前轴总载 = 总重 * 前轴占比；前轴轮数按 (轮数+1)/2 取整，奇数轮时前轴多分 1 个轮。
      单轮载荷 = 前轴总载 / 前轴轮数；轮数不足 2 个或轴距为零时判无效。
  ============================================================
*)
FUNCTION FC_DL_SkateWheelLoadCalc : BOOL
VAR_INPUT
    bEnable      : BOOL; // 使能：TRUE 时计算 / Enable: TRUE to compute
    bErr         : BOOL; // 外部故障：TRUE 时立即退出并置结果无效 / External fault: TRUE aborts with invalid result
    rTotalKg     : REAL; // 滑板与载荷总质量 [kg] / total mass of the skate and the load [kilogram]
    iWheelCnt    : INT;  // 滑板轮总数量 [个] / total number of skate wheels [unit]
    rCgOffset_mm : REAL; // 重心相对几何中心的前向偏移 [mm] / forward offset of the centre of gravity from the geometric centre [millimetre]
    rWheelBase_mm : REAL; // 前后轴距 [mm] / distance between the front and rear axles [millimetre]
END_VAR
VAR_OUTPUT
    rFrontShare : REAL; // 前轴载荷占比，限幅 0.1~0.9 [无量纲] / front axle load share clamped to 0.1 to 0.9 [dimensionless]
    rFrontKg    : REAL; // 前轴总载荷 [kg] / total load on the front axle [kilogram]
    iFrontWheelCnt : INT; // 前轴轮数量 [个] / number of wheels on the front axle [unit]
    rPerWheelKg : REAL; // 前轴单个轮的平均载荷 [kg] / average load of one front wheel [kilogram]
    bValid      : BOOL; // 输出有效：TRUE 表示结果可用 / Output valid
END_VAR
VAR CONSTANT
    DL_R_MAX    : REAL := 3.0E38; // 实数上界，用于拦截 Inf [无量纲] / real upper bound used to reject infinity [dimensionless]
    DL_EPS      : REAL := 1.0E-12; // 除零判定阈值 [无量纲] / division guard threshold [dimensionless]
    DL_HALF     : REAL := 0.5;    // 二分之一，均分基准占比 [无量纲] / one half, the balanced share baseline [dimensionless]
    DL_SHARE_LO : REAL := 0.1;    // 前轴占比下限 [无量纲] / lower clamp of the front share [dimensionless]
    DL_SHARE_HI : REAL := 0.9;    // 前轴占比上限 [无量纲] / upper clamp of the front share [dimensionless]
    DL_WHEEL_MIN : INT := 2;      // 轮数下界 [个] / lower bound of the wheel count [unit]
    DL_WHEEL_MAX : INT := 32;     // 轮数上界 [个] / upper bound of the wheel count [unit]
    DL_BASE_MAX : REAL := 10000.0; // 轴距合理上限 [mm] / sanity upper bound of the wheel base [millimetre]
    DL_MASS_MAX : REAL := 100000.0; // 总质量合理上限 [kg] / sanity upper bound of the total mass [kilogram]
    DL_TWO      : INT := 2;       // 取半数用的除数 [无量纲] / divisor used to obtain half of the wheel count [dimensionless]
    DL_ONE      : INT := 1;       // 奇数轮进位偏置 [个] / carry bias used for an odd wheel count [unit]
END_VAR
VAR
    _bFin    : BOOL := FALSE; // 输入有限性判定结果 / input finiteness verdict
    _rShare  : REAL := 0.0;   // 限幅前前轴占比 [无量纲] / raw front share before clamping [dimensionless]
    _rFrontW : REAL := 0.0;   // 前轴轮数折算实数 [个] / front wheel count cast to real [unit]
END_VAR

    // 段 1｜出口预置：占比先置均分，避免下游误用零
    rFrontShare := DL_HALF;
    rFrontKg := 0.0;
    iFrontWheelCnt := 0;
    rPerWheelKg := 0.0;
    bValid := FALSE;
    // 段 2｜使能闸与外部故障闸
    IF NOT bEnable THEN
        RETURN;
    END_IF;
    IF bErr THEN
        RETURN;
    END_IF;
    // 段 3｜非有限闸
    _bFin := (rTotalKg = rTotalKg) AND (ABS(rTotalKg) <= DL_R_MAX) AND (rCgOffset_mm = rCgOffset_mm) AND (ABS(rCgOffset_mm) <= DL_R_MAX) AND (rWheelBase_mm = rWheelBase_mm) AND (ABS(rWheelBase_mm) <= DL_R_MAX);
    IF NOT _bFin THEN
        RETURN;
    END_IF;
    // 段 4｜域闸：轴距严格为正且合理，总质量非负且合理，轮数 2~32
    IF (ABS(rWheelBase_mm) <= DL_EPS) OR (rWheelBase_mm < 0.0) OR (rWheelBase_mm > DL_BASE_MAX) THEN
        RETURN;
    END_IF;
    IF (rTotalKg < 0.0) OR (rTotalKg > DL_MASS_MAX) THEN
        RETURN;
    END_IF;
    IF (iWheelCnt < DL_WHEEL_MIN) OR (iWheelCnt > DL_WHEEL_MAX) THEN
        RETURN;
    END_IF;
    // 段 5｜前轴占比与限幅
    _rShare := DL_HALF + rCgOffset_mm / rWheelBase_mm;
    IF _rShare < DL_SHARE_LO THEN
        rFrontShare := DL_SHARE_LO;
    ELSIF _rShare > DL_SHARE_HI THEN
        rFrontShare := DL_SHARE_HI;
    ELSE
        rFrontShare := _rShare;
    END_IF;
    // 段 6｜前轴轮数：奇数轮时前轴多分一个
    iFrontWheelCnt := (iWheelCnt + DL_ONE) / DL_TWO;
    IF iFrontWheelCnt < DL_ONE THEN
        iFrontWheelCnt := DL_ONE;
    END_IF;
    // 段 7｜前轴总载与单轮载荷
    rFrontKg := rTotalKg * rFrontShare;
    _rFrontW := INT_TO_REAL(iFrontWheelCnt);
    IF ABS(_rFrontW) <= DL_EPS THEN
        RETURN;
    END_IF;
    rPerWheelKg := rFrontKg / _rFrontW;
    bValid := TRUE;
    FC_DL_SkateWheelLoadCalc := bValid;
END_FUNCTION
